(* CODESYS project beveling.project

Project tree, tasks and I/O mapping:
  Device : AM523-0808TN, Shenzhen Inovance Control Technology, version 3.5.11.50
      settings: PersistentStartAdddr = 0; PersistentStartEndAddr = 524287; Mode = 1
    application Application
      libraries: Standard, * (System); CmpEventMgr, 3.5.8.0 (System); Component Manager, 3.5.9.0 (System); CmpApp, 3.5.11.0 (System); CmpIecTask, 3.5.9.0 (System)
      task MainTask (cyclic, interval 4 ms, priority 1) calls nothing
      task ETHERCAT1 (cyclic, interval 2000 µs, priority 0) calls ETHERCAT1.EtherCAT_Task, PLC_PRG
      90_Legacy/
        program PRG_AxisDemo [ST]
      00_Types/
        data type ST_DeviceConfig
        data type ST_DeviceStatus
        data type E_AutoStep
        data type ST_ManualCommand
        data type ST_SimulationSettings
        data type ST_Recipe
        data type ST_DeviceCommand
        data type E_DeviceAction
        data type E_MachineState
        data type ST_OperatorCommand
        data type E_MachineMode
        data type ST_MachineStatus
        data type E_DeviceKind
      01_Data/
        global variables GVL_Simulation
        global variables GVL_Interface
        global variables GVL_IO
        global variables GVL_Modbus
        global variables GVL_Parameters
        global variables GVL_DeviceIds
      05_Communication/
        function block FB_ModbusInterface [ST]
      06_Simulation/
        function block FB_SimDevice [ST]
        function block FB_SimPlant [ST]
      global variables GVL_Motion
      DifferentialMonitor
      03_Units/
        function block FB_ResetLength [ST]
        function block FB_Unload [ST]
        function block FB_ClearLength [ST]
        function block FB_Initialize [ST]
        function block FB_ClearanceUnit [ST]
        function block FB_ReturnKnife [ST]
        function block FB_ClearTransfer [ST]
        function block FB_PostCut [ST]
      04_Machine/
        function F_RecipeValid [ST]
        function block FB_IOMap [ST]
        function block FB_Machine [ST]
        function block FB_AutoCycle [ST]
        function block FB_Interlocks [ST]
        function block FB_AlarmManager [ST]
        function block FB_ManualControl [ST]
      02_Devices/
        function block FB_Motor [ST]
        function F_At [ST]
        function block FB_Axis [ST]
        function block FB_DeviceManager [ST]
        function F_NextID [ST]
        function F_Done [ST]
        function block FB_Valve [ST]
        function F_Command [ST]
        function block FB_Cylinder [ST]
      program PLC_PRG [ST]
      TaskEventPreStart
    HardWare Configuration
    Network Configuration
      EtherCAT Config
      LocalBus Config
    Resources List
    ConfigStorage
    Device Diagnosis
    HwConfiguratioinDevice : SystemConfig, Inovance, version 00.00.00.10
        settings: NetworkConfigArray.NetworkConfigArray.BusType = 10; NetworkConfigArray.NetworkConfigArray.RackSum = 1; NetworkConfigArray.NetworkConfigArray.HardwareConfigArray.HardwareConfigArray.RackNo = 1
    EXP_A : 扩展卡, 汇川技术股份有限公司, version 00.00.00.10
    ETHERCAT1 : EtherCAT Master SoftMotion, 3S - Smart Software Solutions GmbH, version 3.5.11.10
        settings:  = 0; MasterCycleTime = 2000; NetworkName = 'eth1'; SelectNetworkByName = TRUE; DisableTaskGeneration = True; SlaveArrayName = ADR(_EC1_Node)
      InoSV660N : SV660_1Axis_00915, Inovance, order no. InoSV660N, version Revision=16#00010000
          settings: Number of Outputs = 6; Number of Inputs = 10; Number of Infos about Outputs = 6; Number of Infos about Inputs = 10; Configuration address of the slave = 1; Sync.Length = 18; Sync.Length = 32; FMMU.Length = 18; FMMU.Length = 32; DC sync0 cycletime = 2000; DC sync1 cycletime = 2000; Number of SDO = 10; Homing method.Index = 16#6098; Homing method.Subindex = 16#00; Homing method.Value = 1; Homing method.Size = 8; Homing method.AbortIfError = FALSE; Homing method.JumpToLine = FALSE; Homing method.Line = 0; Homing method.CompleteAccess = FALSE; Actual Position Calculation Method.Index = 16#60E6; Actual Position Calculation Method.Subindex = 16#00; Actual Position Calculation Method.Value = 0; Actual Position Calculation Method.Size = 8; Actual Position Calculation Method.AbortIfError = FALSE; Actual Position Calculation Method.JumpToLine = FALSE; Actual Position Calculation Method.Line = 0; Actual Position Calculation Method.CompleteAccess = FALSE; Speed during search for switch.Index = 16#6099; Speed during search for switch.Subindex = 16#01; Speed during search for switch.Value = 1398102; Speed during search for switch.Size = 32; Speed during search for switch.AbortIfError = FALSE; Speed during search for switch.JumpToLine = FALSE; Speed during search for switch.Line = 0; Speed during search for switch.CompleteAccess = FALSE; Homing acceleration.Index = 16#609A; Homing acceleration.Subindex = 16#00; Homing acceleration.Value = 139810133; Homing acceleration.Size = 32;
            Homing acceleration.AbortIfError = FALSE; Homing acceleration.JumpToLine = FALSE; Homing acceleration.Line = 0; Homing acceleration.CompleteAccess = FALSE; Speed during search for zero.Index = 16#6099; Speed during search for zero.Subindex = 16#02; Speed during search for zero.Value = 139810; Speed during search for zero.Size = 32; Speed during search for zero.AbortIfError = FALSE; Speed during search for zero.JumpToLine = FALSE; Speed during search for zero.Line = 0; Speed during search for zero.CompleteAccess = FALSE; Time of home searching.Index = 16#2005; Time of home searching.Subindex = 16#24; Time of home searching.Value = 50000; Time of home searching.Size = 16; Time of home searching.AbortIfError = FALSE; Time of home searching.JumpToLine = FALSE; Time of home searching.Line = 0; Time of home searching.CompleteAccess = FALSE; Positive torque limit value.Index = 16#60E0; Positive torque limit value.Subindex = 16#00; Positive torque limit value.Value = 3500; Positive torque limit value.Size = 16; Positive torque limit value.AbortIfError = FALSE; Positive torque limit value.JumpToLine = FALSE; Positive torque limit value.Line = 0; Positive torque limit value.CompleteAccess = FALSE; Negative torque limit value.Index = 16#60E1; Negative torque limit value.Subindex = 16#00; Negative torque limit value.Value = 3500; Negative torque limit value.Size = 16; Negative torque limit value.AbortIfError = FALSE; Negative torque limit value.JumpToLine = FALSE; Negative torque limit value.Line = 0; Negative torque limit value.CompleteAccess = FALSE; Max profile velocity.Index = 16#607F; Max profile velocity.Subindex = 16#00; Max profile velocity.Value = 83886080; Max profile velocity.Size = 32;
            Max profile velocity.AbortIfError = FALSE; Max profile velocity.JumpToLine = FALSE; Max profile velocity.Line = 0; Max profile velocity.CompleteAccess = FALSE; RxTxPdo.NumberofEntries = 6; RxTxPdo.Sm = 2; Controlword.Index = 16#6040; Controlword.SubIndex = 0; Controlword.Size = 16; Controlword.DependOnSlot = false; Controlword.DependOnSlotGroup = false; Target position.Index = 16#607A; Target position.SubIndex = 0; Target position.Size = 32; Target position.DependOnSlot = false; Target position.DependOnSlotGroup = false; Touch probe function.Index = 16#60B8; Touch probe function.SubIndex = 0; Touch probe function.Size = 16; Touch probe function.DependOnSlot = false; Touch probe function.DependOnSlotGroup = false; Physical outputs.Index = 16#60FE; Physical outputs.SubIndex = 1; Physical outputs.Size = 32; Physical outputs.DependOnSlot = false; Physical outputs.DependOnSlotGroup = false; Target velocity.Index = 16#60FF; Target velocity.SubIndex = 0; Target velocity.Size = 32; Target velocity.DependOnSlot = false; Target velocity.DependOnSlotGroup = false; Target torque.Index = 16#6071; Target torque.SubIndex = 0; Target torque.Size = 16; Target torque.DependOnSlot = false; Target torque.DependOnSlotGroup = false; RxTxPdo.Sm = -1; RxTxPdo.NumberofEntries = 10; RxTxPdo.Sm = 3; Error code.Index = 16#603F;
            Error code.SubIndex = 0; Error code.Size = 16; Error code.DependOnSlot = false; Error code.DependOnSlotGroup = false; Statusword.Index = 16#6041; Statusword.SubIndex = 0; Statusword.Size = 16; Statusword.DependOnSlot = false; Statusword.DependOnSlotGroup = false; Position actual value.Index = 16#6064; Position actual value.SubIndex = 0; Position actual value.Size = 32; Position actual value.DependOnSlot = false; Position actual value.DependOnSlotGroup = false; Torque actual value.Index = 16#6077; Torque actual value.SubIndex = 0; Torque actual value.Size = 16; Torque actual value.DependOnSlot = false; Torque actual value.DependOnSlotGroup = false; Following error actual value.Index = 16#60F4; Following error actual value.SubIndex = 0; Following error actual value.Size = 32; Following error actual value.DependOnSlot = false; Following error actual value.DependOnSlotGroup = false; Touch probe status.Index = 16#60B9; Touch probe status.SubIndex = 0; Touch probe status.Size = 16; Touch probe status.DependOnSlot = false; Touch probe status.DependOnSlotGroup = false; Touch probe pos1 pos value.Index = 16#60BA; Touch probe pos1 pos value.SubIndex = 0; Touch probe pos1 pos value.Size = 32; Touch probe pos1 pos value.DependOnSlot = false; Touch probe pos1 pos value.DependOnSlotGroup = false; Touch probe pos2 pos value.Index = 16#60BC; Touch probe pos2 pos value.SubIndex = 0; Touch probe pos2 pos value.Size = 32; Touch probe pos2 pos value.DependOnSlot = false; Touch probe pos2 pos value.DependOnSlotGroup = false; Digital inputs.Index = 16#60FD;
            Digital inputs.SubIndex = 0; Digital inputs.Size = 32; Digital inputs.DependOnSlot = false; Digital inputs.DependOnSlotGroup = false; Velocity actual value.Index = 16#606C; Velocity actual value.SubIndex = 0; Velocity actual value.Size = 32; Velocity actual value.DependOnSlot = false; Velocity actual value.DependOnSlotGroup = false; RxTxPdo.Sm = -1; Controlword.Name = 'Controlword'; Controlword.DataType = 'UINT'; Target position.Name = 'Target position'; Target position.DataType = 'DINT'; Touch probe function.Name = 'Touch probe function'; Touch probe function.DataType = 'UINT'; Physical outputs.Name = 'Physical outputs'; Physical outputs.DataType = 'UDINT'; Target velocity.Name = 'Target velocity'; Target velocity.DataType = 'DINT'; Target torque.Name = 'Target torque'; Target torque.DataType = 'INT'; Error code.Name = 'Error code'; Error code.DataType = 'UINT'; Statusword.Name = 'Statusword'; Statusword.DataType = 'UINT'; Position actual value.Name = 'Position actual value'; Position actual value.DataType = 'DINT'; Torque actual value.Name = 'Torque actual value'; Torque actual value.DataType = 'INT'; Following error actual value.Name = 'Following error actual value'; Following error actual value.DataType = 'DINT'; Touch probe status.Name = 'Touch probe status'; Touch probe status.DataType = 'UINT'; Touch probe pos1 pos value.Name = 'Touch probe pos1 pos value'; Touch probe pos1 pos value.DataType = 'DINT'; Touch probe pos2 pos value.Name = 'Touch probe pos2 pos value'; Touch probe pos2 pos value.DataType = 'DINT'; Digital inputs.Name = 'Digital inputs'; Digital inputs.DataType = 'UDINT';
            Velocity actual value.Name = 'Velocity actual value'; Velocity actual value.DataType = 'DINT'
          unmapped channels: Controlword, Target position, Touch probe function, Physical outputs, Target velocity, Target torque, Error code, Statusword, Position actual value, Torque actual value, Following error actual value, Touch probe status, Touch probe pos1 pos value, Touch probe pos2 pos value, Digital inputs, Velocity actual value
        Axis_1 : Axis, 3S - Smart Software Solutions GmbH, order no. 0, version 4.0.0.0
            settings: wDriveID = 0; dwRatioTechUnitsDenom = 4194304; iRatioTechUnitsNum = 5; HomingMode = 10; ZeroSignal = 0; StartDirction = 1; EndDirection = 1; PosLimitMode = 0; NegLimitMode = 0; HomingVelocity = 10; HomingApproachVelocity = 2; HomingAcceleration = 100; HomingDeceleration = 100; HomingJerk = 0; HomeMaskDistance = 0; HomePositionOffset = 0; HomePushTime = 0; HomeCompensation = 0; HomeTimeout = 0; HomeCompensationVelocity = 1000; 4000 = 1; 4001 = 0; 4003 = true; 4004 = 3; 4005 = 0; 4006 = 1.666667; 4007 = 166.666666; 4008 = 0.166667; 4009 = 50000; 4010 = 3500; 4011 = 3500; 4012 = 100.000000; ScalingIncs = 16#800000; 6005 = 10; AdrOffset_8010 = 4; BitOffset_8010 = 0; BitLength_8010 = 16; Address_8010 = '%QW2'; Type_8010 = 'UINT'; AddressPointer_8010 = ADR(%QW2);
              AdrOffset_8020 = 8; BitOffset_8020 = 0; BitLength_8020 = 32; Address_8020 = '%QD2'; Type_8020 = 'DINT'; AddressPointer_8020 = ADR(%QD2); AdrOffset_8030 = 20; BitOffset_8030 = 0; BitLength_8030 = 32; Address_8030 = '%QD5'; Type_8030 = 'DINT'; AddressPointer_8030 = ADR(%QD5); AdrOffset_8040 = 24; BitOffset_8040 = 0; BitLength_8040 = 16; Address_8040 = '%QW12'; Type_8040 = 'INT'; AddressPointer_8040 = ADR(%QW12); AdrOffset_8050 = 4294967295; BitOffset_8050 = 0; BitLength_8050 = 0; Address_8050 = ''; Type_8050 = ''; AddressPointer_8050 = 0; AdrOffset_8060 = 12; BitOffset_8060 = 0; BitLength_8060 = 16; Address_8060 = '%QW6'; Type_8060 = 'UINT'; AddressPointer_8060 = ADR(%QW6); AdrOffset_8070 = 4294967295; BitOffset_8070 = 0; BitLength_8070 = 0; Address_8070 = ''; Type_8070 = ''; AddressPointer_8070 = 0; AdrOffset_8080 = 4294967295; BitOffset_8080 = 0; BitLength_8080 = 0; Address_8080 = '';
              Type_8080 = ''; AddressPointer_8080 = 0; AdrOffset_8090 = 16; BitOffset_8090 = 0; BitLength_8090 = 32; Address_8090 = '%QD4'; Type_8090 = 'UDINT'; AddressPointer_8090 = ADR(%QD4); AdrOffset_8100 = 4294967295; BitOffset_8100 = 0; BitLength_8100 = 0; Address_8100 = ''; Type_8100 = ''; AddressPointer_8100 = 0; AdrOffset_8510 = 6; BitOffset_8510 = 0; BitLength_8510 = 16; Address_8510 = '%IW3'; Type_8510 = 'UINT'; AddressPointer_8510 = ADR(%IW3); AdrOffset_8520 = 8; BitOffset_8520 = 0; BitLength_8520 = 32; Address_8520 = '%ID2'; Type_8520 = 'DINT'; AddressPointer_8520 = ADR(%ID2); AdrOffset_8530 = 36; BitOffset_8530 = 0; BitLength_8530 = 32; Address_8530 = '%ID9'; Type_8530 = 'DINT'; AddressPointer_8530 = ADR(%ID9); AdrOffset_8540 = 12; BitOffset_8540 = 0; BitLength_8540 = 16; Address_8540 = '%IW6'; Type_8540 = 'INT'; AddressPointer_8540 = ADR(%IW6); AdrOffset_8550 = 4294967295; BitOffset_8550 = 0;
              BitLength_8550 = 0; Address_8550 = ''; Type_8550 = ''; AddressPointer_8550 = 0; AdrOffset_8560 = 32; BitOffset_8560 = 0; BitLength_8560 = 32; Address_8560 = '%ID8'; Type_8560 = 'UDINT'; AddressPointer_8560 = ADR(%ID8); AdrOffset_8570 = 20; BitOffset_8570 = 0; BitLength_8570 = 16; Address_8570 = '%IW10'; Type_8570 = 'UINT'; AddressPointer_8570 = ADR(%IW10); AdrOffset_8580 = 24; BitOffset_8580 = 0; BitLength_8580 = 32; Address_8580 = '%ID6'; Type_8580 = 'DINT'; AddressPointer_8580 = ADR(%ID6); AdrOffset_8590 = 4294967295; BitOffset_8590 = 0; BitLength_8590 = 0; Address_8590 = ''; Type_8590 = ''; AddressPointer_8590 = 0; AdrOffset_8600 = 28; BitOffset_8600 = 0; BitLength_8600 = 32; Address_8600 = '%ID7'; Type_8600 = 'DINT'; AddressPointer_8600 = ADR(%ID7); AdrOffset_8600 = 4294967295; BitOffset_8600 = 0; BitLength_8600 = 0; Address_8610 = ''; Type_8610 = ''; AddressPointer_8610 = 0;
              AdrOffset_8620 = 4; BitOffset_8620 = 0; BitLength_8620 = 16; Address_8620 = '%IW2'; Type_8620 = 'UINT'; AddressPointer_8620 = ADR(%IW2); IsValid = True; AxisNumber = 1; IsHostHoming = True; PulseSelectIndex = 4; SERVO_MAX_ID = 83886080
    SoftMotion General Axis Pool
    Serial : 串行接口, 汇川技术股份有限公司, version 00.00.00.10
      COM : Serial Port, Inovance, version 00.00.00.10
          settings: Device = AM523-0808TN; devGuid = 'e48f0cf2-85a4-455f-a8e7-135d3403221f'
    Local Bus
    EXP_B : 扩展卡, 汇川技术股份有限公司, version 00.00.00.10
    MODBUS_TCP : ModbusTCP本地从站, inovance, version 00.00.00.10
    LocalHSIO : 本地高速IO, 汇川技术股份有限公司, version 2.0.0.0
        unmapped channels: DigitalInput, DigitalOutput
    CAN : CAN总线, INOVANCE, version 00.00.00.10
*)

// Device/Application/00_Types/ST_DeviceConfig
TYPE ST_DeviceConfig :
STRUCT
eKind : E_DeviceKind;
lrInitialPosition : LREAL;
lrMinPosition : LREAL := -1000.0;
lrMaxPosition : LREAL := 1000.0;
lrMaxVelocity : LREAL := 100.0;
tSimAction : TIME := T#500MS;
END_STRUCT
END_TYPE

// Device/Application/00_Types/ST_DeviceStatus
TYPE ST_DeviceStatus :
STRUCT
xReady : BOOL;
xBusy : BOOL;
xActive : BOOL;
xError : BOOL;
udiErrorID : UDINT;
udiAcceptedID : UDINT;
udiCompletedID : UDINT;
lrPosition : LREAL;
END_STRUCT
END_TYPE

// Device/Application/00_Types/E_AutoStep
{attribute 'qualified_only'}
TYPE E_AutoStep :
(
    Idle := 0,
    FeedWait := 10,
    StopFeed := 20,
    Push := 30,
    Clearance := 40,
    Rotate := 50,
    PressDown := 60,
    KnifeDown := 70,
    SpindleOn := 80,
    Cutting := 90,
    StopCut := 100,
    PostCut := 110,
    Complete := 120,
    Fault := 900
);
END_TYPE

// Device/Application/00_Types/ST_ManualCommand
TYPE ST_ManualCommand :
STRUCT
xJogPositive : BOOL;
xJogNegative : BOOL;
xMove : BOOL;
xRun : BOOL;
lrTarget : LREAL;
lrVelocity : LREAL := 10.0;
END_STRUCT
END_TYPE

// Device/Application/00_Types/ST_SimulationSettings
TYPE ST_SimulationSettings :
STRUCT
xSafetyOK : BOOL := TRUE;
xAutoMaterial : BOOL := TRUE;
xMaterialSensor : BOOL;
tMaterialDelay : TIME := T#1S;
axStall : ARRAY[1..17] OF BOOL;
axFault : ARRAY[1..17] OF BOOL;
END_STRUCT
END_TYPE

// Device/Application/00_Types/ST_Recipe
TYPE ST_Recipe :
STRUCT
uiMaterialModel : UINT := 300;
lrCutHome : LREAL := 0.0;
lrCutLength : LREAL := 20.0;
lrCutVelocity : LREAL := 10.0;
lrPositionVelocity : LREAL := 10.0;
lrBeltVelocity : LREAL := 10.0;
lrSpindleVelocity : LREAL := 10.0;
lrLengthPosition : LREAL := 100.0;
lrLengthClear : LREAL := 0.0;
lrRotateAngle : LREAL := 0.0;
lrGripperFront : LREAL := 100.0;
lrGripperPull : LREAL := 200.0;
lrGripperBack : LREAL := 50.0;
lrGripperHome : LREAL := 0.0;
tSpray : TIME := T#300MS;
tStepTimeout : TIME := T#30S;
END_STRUCT
END_TYPE

// Device/Application/00_Types/ST_DeviceCommand
TYPE ST_DeviceCommand :
STRUCT
eAction : E_DeviceAction;
udiID : UDINT;
lrTarget : LREAL;
lrVelocity : LREAL;
END_STRUCT
END_TYPE

// Device/Application/00_Types/E_DeviceAction
{attribute 'qualified_only'}
TYPE E_DeviceAction :
(
    None := 0,
    Position := 1,
    Run := 2,
    Jog := 3,
    Stop := 4
);
END_TYPE

// Device/Application/00_Types/E_MachineState
{attribute 'qualified_only'}
TYPE E_MachineState :
(
    Stopped := 0,
    Initializing := 10,
    Ready := 20,
    Manual := 30,
    Automatic := 40,
    Fault := 90
);
END_TYPE

// Device/Application/00_Types/ST_OperatorCommand
TYPE ST_OperatorCommand :
STRUCT
eMode : E_MachineMode := E_MachineMode.Manual;
xInitialize : BOOL;
xStart : BOOL;
xStop : BOOL;
xResetAlarm : BOOL;
xContinuous : BOOL;
xRemoteControl : BOOL;
END_STRUCT
END_TYPE

// Device/Application/00_Types/E_MachineMode
{attribute 'qualified_only'}
TYPE E_MachineMode :
(
    Manual := 0,
    Automatic := 1
);
END_TYPE

// Device/Application/00_Types/ST_MachineStatus
TYPE ST_MachineStatus :
STRUCT
eState : E_MachineState;
eMode : E_MachineMode;
eAutoStep : E_AutoStep;
xSimulation : BOOL;
xRealBackendAvailable : BOOL;
xInitialized : BOOL;
xReady : BOOL;
xMaterialAtLength : BOOL;
xCycleComplete : BOOL;
udiCycleCount : UDINT;
udiAlarm : UDINT;
uiBlockedDevice : UINT;
uiManualReject : UINT;
uiClearLengthStep : UINT;
uiClearTransferStep : UINT;
uiPostStep : UINT;
uiReturnKnifeStep : UINT;
uiUnloadStep : UINT;
uiResetLengthStep : UINT;
uiInitializeStep : UINT;
uiActiveMaterialModel : UINT;
wRemoteAckSequence : WORD;
uiRemoteResult : UINT;
END_STRUCT
END_TYPE

// Device/Application/00_Types/E_DeviceKind
{attribute 'qualified_only'}
TYPE E_DeviceKind :
(
    Unused := 0,
    Axis := 1,
    Motor := 2,
    Cylinder := 3,
    Valve := 4
);
END_TYPE

// Device/Application/01_Data/GVL_Simulation
VAR_GLOBAL
    stSettings : ST_SimulationSettings;
END_VAR

// Device/Application/01_Data/GVL_Interface
VAR_GLOBAL
    stPanel : ST_OperatorCommand;
    aManual : ARRAY[1..17] OF ST_ManualCommand;
    stStatus : ST_MachineStatus;
    aDeviceStatus : ARRAY[1..17] OF ST_DeviceStatus;
END_VAR

// Device/Application/01_Data/GVL_IO
VAR_GLOBAL
    (* Unmapped interface. No AT %Q / %I bindings in this framework. *)
    xSafetyOK : BOOL;
    xMaterialAtLength : BOOL;
    axDigitalInputs : ARRAY[0..31] OF BOOL;
    axDigitalOutputs : ARRAY[0..31] OF BOOL;
    axG2RelayDemand : ARRAY[1..3] OF BOOL;
END_VAR

// Device/Application/01_Data/GVL_Modbus
VAR_GLOBAL
    (* Buffers only; the existing MODBUS_TCP driver is not bound yet. *)
    xEnable : BOOL;
    awRx : ARRAY[0..31] OF WORD;
    awTx : ARRAY[0..127] OF WORD;
END_VAR

// Device/Application/GVL_Motion
VAR_GLOBAL
    (* ================= Commands (HMI / online write) ================= *)
    xEnable     : BOOL;              (* power on / off the servo axis *)
    xReset      : BOOL;              (* reset axis error *)
    xStop       : BOOL;              (* stop and lock the axis *)
    xJogFwd     : BOOL;              (* jog forward (level) *)
    xJogRev     : BOOL;              (* jog reverse (level) *)
    xMoveRel    : BOOL;              (* relative move command (level) *)
    xMoveAbs    : BOOL;              (* absolute move command (level) *)
    xStartCycle : BOOL;              (* start auto fwd/back cycle (rising edge) *)

    rRelDist    : LREAL := 100.0;    (* relative move distance [mm] *)
    rTargetPos  : LREAL := 0.0;      (* absolute target position [mm] *)

    (* ================= Motion parameters ================= *)
    rJogVel     : LREAL := 10.0;     (* jog velocity [mm/s] *)
    rVel        : LREAL := 30.0;     (* positioning velocity [mm/s] *)
    rAcc        : LREAL := 200.0;    (* acceleration [mm/s2] *)
    rDec        : LREAL := 200.0;    (* deceleration [mm/s2] *)
    rStroke     : LREAL := 100.0;    (* auto cycle stroke (one way) [mm] *)
    tDwell      : TIME  := T#1S;     (* dwell time at cycle ends *)

    (* ================= Status ================= *)
    xPowered    : BOOL;              (* MC_Power.Status : servo enabled *)
    xAxisReady  : BOOL;              (* axis in StandStill -> motion allowed *)
    xBusy       : BOOL;              (* any motion active *)
    xDisabled   : BOOL;              (* axis state = Disabled *)
    xStandStill : BOOL;              (* axis state = StandStill *)
    xStopping   : BOOL;              (* axis state = Stopping *)
    xErrorStop  : BOOL;              (* axis state = ErrorStop *)
    xAxisError  : BOOL;              (* axis reports an error *)
    iAxisErrorID: DWORD;             (* axis error code *)
    rActPos     : LREAL;             (* actual position [mm] *)
    iState      : INT;               (* auto cycle step number *)
END_VAR

// Device/Application/01_Data/GVL_Parameters
VAR_GLOBAL
    (* Simulation examples only: these are NOT commissioned machine settings. *)
    xSimulation : BOOL := TRUE;
    stRecipe : ST_Recipe;
END_VAR

// Device/Application/01_Data/GVL_DeviceIds
VAR_GLOBAL CONSTANT
    D1_Belt : UINT := 1;
    D2_CutFeed : UINT := 2;
    D3_Spindle : UINT := 3;
    D4_LengthMove : UINT := 4;
    D5_LengthLift : UINT := 5;
    D7_GripperMove : UINT := 7;
    D8_Rotate : UINT := 8;
    G1_Press : UINT := 9;
    G2_SideStop : UINT := 10;
    G3_Push : UINT := 11;
    G4_RollerLift : UINT := 12;
    G5_Spray : UINT := 13;
    G6_Air : UINT := 14;
    G7_GripperLift : UINT := 15;
    G8_GripperClamp : UINT := 16;
    G9_KnifeLift : UINT := 17;
END_VAR

// Device/Application/PLC_PRG
PROGRAM PLC_PRG
VAR
    fbCommunication : FB_ModbusInterface;
    fbMachine : FB_Machine;
    fbIO : FB_IOMap;
END_VAR

(* One cyclic owner in ETHERCAT1. All lower device FBs are called each scan. *)
fbCommunication(xEnable:=GVL_Modbus.xEnable,stStatus:=GVL_Interface.stStatus,
    aStatus:=GVL_Interface.aDeviceStatus,awRx:=GVL_Modbus.awRx,awTx:=GVL_Modbus.awTx);
fbMachine(xSimulation:=GVL_Parameters.xSimulation,stPanel:=GVL_Interface.stPanel,
    stRemote:=fbCommunication.stCommand,xRemoteRequest:=fbCommunication.xRequest,
    wRemoteSequence:=fbCommunication.wRequestSequence,aManual:=GVL_Interface.aManual,
    stRecipe:=GVL_Parameters.stRecipe,stSim:=GVL_Simulation.stSettings,
    xRealSafetyOK:=GVL_IO.xSafetyOK,xRealMaterial:=GVL_IO.xMaterialAtLength);
GVL_Interface.stStatus:=fbMachine.stStatus;
GVL_Interface.aDeviceStatus:=fbMachine.aDeviceStatus;
fbIO(uiMaterialModel:=fbMachine.stStatus.uiActiveMaterialModel,aCommand:=fbMachine.aSelectedCommand,
    aStatus:=fbMachine.aDeviceStatus,
    axOutputs:=GVL_IO.axDigitalOutputs,axG2RelayDemand:=GVL_IO.axG2RelayDemand);

END_PROGRAM

// Device/Application/05_Communication/FB_ModbusInterface
FUNCTION_BLOCK FB_ModbusInterface
VAR_INPUT
    xEnable : BOOL;
    stStatus : ST_MachineStatus;
    aStatus : ARRAY[1..17] OF ST_DeviceStatus;
END_VAR
VAR_IN_OUT
    awRx : ARRAY[0..31] OF WORD;
    awTx : ARRAY[0..127] OF WORD;
END_VAR
VAR_OUTPUT
    xRequest : BOOL;
    wRequestSequence : WORD;
    stCommand : ST_OperatorCommand;
    uiParseResult : UINT;
END_VAR
VAR
    aSnapshot : ARRAY[0..31] OF WORD;
    wLastSeen : WORD;
    xWasEnabled : BOOL;
    i : INT;
END_VAR

xRequest:=FALSE;
stCommand.xInitialize:=FALSE; stCommand.xStart:=FALSE;
stCommand.xStop:=FALSE; stCommand.xResetAlarm:=FALSE;
IF NOT xEnable OR NOT xWasEnabled THEN
    (* Baseline on enable, so reconnect never replays a stale command. *)
    wLastSeen:=awRx[1];
ELSIF (awRx[1]<>0) AND (awRx[1]<>wLastSeen) THEN
    aSnapshot:=awRx;
    IF aSnapshot[1]=awRx[1] THEN
        wLastSeen:=aSnapshot[1]; wRequestSequence:=aSnapshot[1]; uiParseResult:=0;
        IF (aSnapshot[0]<>1) OR (aSnapshot[3]>1) OR (aSnapshot[2]<1) OR (aSnapshot[2]>4) THEN
            uiParseResult:=2;
        ELSE
            IF aSnapshot[3]=0 THEN stCommand.eMode:=E_MachineMode.Manual;
            ELSE stCommand.eMode:=E_MachineMode.Automatic; END_IF
            stCommand.xContinuous:=aSnapshot[4]<>0;
            CASE aSnapshot[2] OF
            1: stCommand.xInitialize:=TRUE;
            2: stCommand.xStart:=TRUE;
            3: stCommand.xStop:=TRUE;
            4: stCommand.xResetAlarm:=TRUE;
            END_CASE
            xRequest:=TRUE;
        END_IF
    END_IF
END_IF
xWasEnabled:=xEnable;
FOR i:=0 TO 127 DO awTx[i]:=0; END_FOR
awTx[0]:=1; awTx[1]:=stStatus.wRemoteAckSequence; awTx[2]:=UINT_TO_WORD(stStatus.uiRemoteResult);
awTx[3]:=TO_WORD(stStatus.eState); awTx[4]:=TO_WORD(stStatus.eAutoStep);
awTx[5]:=UDINT_TO_WORD(stStatus.udiAlarm); awTx[6]:=UDINT_TO_WORD(SHR(stStatus.udiAlarm,16));
awTx[7]:=UDINT_TO_WORD(stStatus.udiCycleCount); awTx[8]:=UDINT_TO_WORD(SHR(stStatus.udiCycleCount,16));
awTx[9]:=BOOL_TO_WORD(stStatus.xSimulation); awTx[10]:=BOOL_TO_WORD(stStatus.xInitialized);
awTx[11]:=BOOL_TO_WORD(stStatus.xMaterialAtLength); awTx[12]:=UINT_TO_WORD(stStatus.uiActiveMaterialModel);
awTx[13]:=wRequestSequence; awTx[14]:=UINT_TO_WORD(uiParseResult);
(* Positions at [32..48]: signed INT, 0.1 engineering-unit scaling. *)
FOR i:=1 TO 17 DO awTx[31+i]:=INT_TO_WORD(LREAL_TO_INT(aStatus[i].lrPosition*10.0)); END_FOR

END_FUNCTION_BLOCK

// Device/Application/04_Machine/FB_Machine
FUNCTION_BLOCK FB_Machine
VAR_INPUT
    xSimulation : BOOL;
    stPanel : ST_OperatorCommand;
    stRemote : ST_OperatorCommand;
    xRemoteRequest : BOOL;
    wRemoteSequence : WORD;
    aManual : ARRAY[1..17] OF ST_ManualCommand;
    stRecipe : ST_Recipe;
    stSim : ST_SimulationSettings;
    xRealSafetyOK : BOOL;
    xRealMaterial : BOOL;
END_VAR
VAR_OUTPUT
    stStatus : ST_MachineStatus;
    aDeviceStatus : ARRAY[1..17] OF ST_DeviceStatus;
    aSelectedCommand : ARRAY[1..17] OF ST_DeviceCommand;
END_VAR
VAR
    stCommand : ST_OperatorCommand;
    stActiveRecipe : ST_Recipe;
    aRequest : ARRAY[1..17] OF ST_DeviceCommand;
    stEmpty : ST_DeviceCommand;
    fbDevices : FB_DeviceManager;
    fbManual : FB_ManualControl;
    fbAuto : FB_AutoCycle;
    fbInitialize : FB_Initialize;
    fbInterlocks : FB_Interlocks;
    fbPlant : FB_SimPlant;
    fbAlarm : FB_AlarmManager;
    rtInitialize : R_TRIG;
    rtStart : R_TRIG;
    rtReset : R_TRIG;
    udiCounter : UDINT;
    udiFault : UDINT;
    xSafetyOK : BOOL;
    xMaterial : BOOL;
    xInitialized : BOOL;
    xPermit : BOOL;
    xRemoteAccepted : BOOL;
    xResetDevices : BOOL;
    xLastSimulation : BOOL := TRUE;
    xManualReleased : BOOL;
    xManualArmed : BOOL;
    eActiveMode : E_MachineMode;
    i : INT;
END_VAR

stCommand:=stPanel;
IF stPanel.xRemoteControl THEN
    (* Mode and continuous selection persist between remote command frames. *)
    stCommand.eMode:=stRemote.eMode;
    stCommand.xContinuous:=stRemote.xContinuous;
END_IF
xRemoteAccepted:=FALSE;
IF xRemoteRequest THEN
    stStatus.wRemoteAckSequence:=wRemoteSequence;
    IF stPanel.xRemoteControl THEN
        stCommand:=stRemote;
        (* Local stop always overrides remote control. *)
        stCommand.xStop:=stCommand.xStop OR stPanel.xStop;
        stStatus.uiRemoteResult:=0; xRemoteAccepted:=TRUE;
    ELSE stStatus.uiRemoteResult:=1;
    END_IF
END_IF
rtInitialize(CLK:=stCommand.xInitialize);
rtStart(CLK:=stCommand.xStart);
rtReset(CLK:=stCommand.xResetAlarm);
IF xSimulation THEN xSafetyOK:=stSim.xSafetyOK; xMaterial:=fbPlant.xMaterialAtLength;
ELSE xSafetyOK:=xRealSafetyOK; xMaterial:=xRealMaterial; END_IF
udiFault:=0;
IF NOT xSafetyOK THEN udiFault:=1001; END_IF
IF NOT xSimulation THEN udiFault:=3001; END_IF
IF xSimulation<>xLastSimulation THEN
    stStatus.eState:=E_MachineState.Stopped; xInitialized:=FALSE;
END_IF
xLastSimulation:=xSimulation;
FOR i:=1 TO 17 DO
    IF aDeviceStatus[i].xError THEN udiFault:=10000+INT_TO_UDINT(i); END_IF
    aRequest[i]:=stEmpty;
END_FOR
IF (stStatus.eState=E_MachineState.Automatic) OR (stStatus.eState=E_MachineState.Manual) THEN
    IF stCommand.eMode<>eActiveMode THEN stStatus.eState:=E_MachineState.Stopped; xInitialized:=FALSE; END_IF
END_IF
IF stCommand.xStop THEN stStatus.eState:=E_MachineState.Stopped; xInitialized:=FALSE; END_IF
IF udiFault<>0 THEN stStatus.eState:=E_MachineState.Fault; xInitialized:=FALSE; END_IF
xResetDevices:=rtReset.Q AND xSafetyOK AND xSimulation;
IF xResetDevices THEN
    (* Reset injected/device errors before clearing the machine latch next scan. *)
    udiFault:=0;
    FOR i:=1 TO 17 DO IF stSim.axFault[i] THEN udiFault:=10000+INT_TO_UDINT(i); END_IF END_FOR
END_IF
fbAlarm(udiIncoming:=udiFault,xReset:=xResetDevices);
IF (stStatus.eState=E_MachineState.Fault) AND (fbAlarm.udiLatched=0) AND xResetDevices THEN
    stStatus.eState:=E_MachineState.Stopped;
END_IF
IF fbAlarm.udiLatched<>0 THEN stStatus.eState:=E_MachineState.Fault; END_IF
IF rtInitialize.Q AND NOT stCommand.xStop THEN
    IF (stStatus.eState=E_MachineState.Stopped) AND xSimulation AND xSafetyOK AND F_RecipeValid(stRecipe) THEN
        stActiveRecipe:=stRecipe; stStatus.eState:=E_MachineState.Initializing;
        eActiveMode:=stCommand.eMode; xInitialized:=FALSE;
    ELSIF xRemoteAccepted THEN stStatus.uiRemoteResult:=3;
    END_IF
END_IF
IF stStatus.eState=E_MachineState.Ready THEN
    IF stCommand.eMode=E_MachineMode.Manual THEN
        stStatus.eState:=E_MachineState.Manual; eActiveMode:=E_MachineMode.Manual;
    ELSIF rtStart.Q AND NOT stCommand.xStop THEN
        IF F_RecipeValid(stRecipe) THEN
            stActiveRecipe:=stRecipe; eActiveMode:=E_MachineMode.Automatic;
            stStatus.eState:=E_MachineState.Automatic;
        ELSIF xRemoteAccepted THEN stStatus.uiRemoteResult:=5;
        END_IF
    END_IF
ELSIF (stStatus.eState=E_MachineState.Manual) AND (stCommand.eMode=E_MachineMode.Automatic) THEN
    stStatus.eState:=E_MachineState.Stopped; xInitialized:=FALSE;
END_IF
IF rtStart.Q AND xRemoteAccepted AND (stStatus.eState<>E_MachineState.Automatic) THEN stStatus.uiRemoteResult:=3; END_IF

xManualReleased:=TRUE;
FOR i:=1 TO 17 DO
    IF aManual[i].xJogPositive OR aManual[i].xJogNegative OR aManual[i].xMove OR aManual[i].xRun THEN xManualReleased:=FALSE; END_IF
END_FOR
IF stStatus.eState<>E_MachineState.Manual THEN xManualArmed:=FALSE;
ELSIF xManualReleased THEN xManualArmed:=TRUE;
END_IF
fbInitialize(xExecute:=stStatus.eState=E_MachineState.Initializing,stRecipe:=stActiveRecipe,
    aCommand:=aRequest,aStatus:=aDeviceStatus,udiCounter:=udiCounter);
fbManual(xEnable:=(stStatus.eState=E_MachineState.Manual) AND xManualArmed,
    aManual:=aManual,aCommand:=aRequest,aStatus:=aDeviceStatus,udiCounter:=udiCounter);
fbAuto(xRun:=stStatus.eState=E_MachineState.Automatic,xContinuous:=stCommand.xContinuous,
    xMaterialAtLength:=xMaterial,stRecipe:=stActiveRecipe,aCommand:=aRequest,aStatus:=aDeviceStatus,udiCounter:=udiCounter);
IF fbInitialize.xDone THEN xInitialized:=TRUE; stStatus.eState:=E_MachineState.Ready; END_IF
IF fbInitialize.xError OR fbAuto.xError THEN
    udiFault:=MAX(fbInitialize.udiErrorID,fbAuto.udiErrorID);
    fbAlarm(udiIncoming:=udiFault,xReset:=FALSE);
    stStatus.eState:=E_MachineState.Fault; xInitialized:=FALSE;
END_IF
IF fbAuto.xDone THEN
    stStatus.udiCycleCount:=stStatus.udiCycleCount+1;
    IF NOT stCommand.xContinuous THEN stStatus.eState:=E_MachineState.Ready; END_IF
END_IF
xPermit:=xSimulation AND xSafetyOK AND NOT stCommand.xStop AND (fbAlarm.udiLatched=0)
    AND ((stStatus.eState=E_MachineState.Initializing) OR (stStatus.eState=E_MachineState.Manual)
    OR (stStatus.eState=E_MachineState.Automatic));
fbInterlocks(xPermit:=xPermit,stRecipe:=stActiveRecipe,aRequest:=aRequest,aStatus:=aDeviceStatus);
aSelectedCommand:=fbInterlocks.aCommand;
fbDevices(xEnable:=xSimulation AND xSafetyOK,xSimulation:=xSimulation,xReset:=xResetDevices,
    stSim:=stSim,aCommand:=aSelectedCommand);
aDeviceStatus:=fbDevices.aStatus;
fbPlant(xEnable:=xSimulation,stSettings:=stSim,aStatus:=aDeviceStatus);
stStatus.eMode:=stCommand.eMode; stStatus.eAutoStep:=fbAuto.eStep;
stStatus.xSimulation:=xSimulation; stStatus.xRealBackendAvailable:=FALSE;
stStatus.xInitialized:=xInitialized;
stStatus.xReady:=xInitialized AND (stStatus.eState=E_MachineState.Ready);
stStatus.xMaterialAtLength:=xMaterial; stStatus.xCycleComplete:=fbAuto.xDone;
stStatus.udiAlarm:=fbAlarm.udiLatched; stStatus.uiBlockedDevice:=fbInterlocks.uiBlockedDevice;
stStatus.uiManualReject:=fbManual.uiRejectDevice;
stStatus.uiClearLengthStep:=fbAuto.uiClearLengthStep; stStatus.uiClearTransferStep:=fbAuto.uiClearTransferStep;
stStatus.uiPostStep:=fbAuto.uiPostStep; stStatus.uiReturnKnifeStep:=fbAuto.uiReturnKnifeStep;
stStatus.uiUnloadStep:=fbAuto.uiUnloadStep; stStatus.uiResetLengthStep:=fbAuto.uiResetLengthStep;
stStatus.uiInitializeStep:=fbInitialize.uiStep; stStatus.uiActiveMaterialModel:=stActiveRecipe.uiMaterialModel;

END_FUNCTION_BLOCK

// Device/Application/04_Machine/F_RecipeValid
FUNCTION F_RecipeValid : BOOL
VAR_INPUT
    stRecipe : ST_Recipe;
END_VAR

F_RecipeValid := ((stRecipe.uiMaterialModel = 300) OR
    (stRecipe.uiMaterialModel = 400) OR (stRecipe.uiMaterialModel = 600))
    AND (stRecipe.lrCutLength > 0.0) AND (stRecipe.lrCutLength <= 500.0)
    AND (stRecipe.lrCutVelocity > 0.0) AND (stRecipe.lrCutVelocity <= 100.0)
    AND (stRecipe.lrPositionVelocity > 0.0) AND (stRecipe.lrPositionVelocity <= 100.0)
    AND (stRecipe.lrBeltVelocity > 0.0) AND (stRecipe.lrBeltVelocity <= 100.0)
    AND (stRecipe.lrSpindleVelocity > 0.0) AND (stRecipe.lrSpindleVelocity <= 100.0)
    AND (stRecipe.tStepTimeout >= T#1S) AND (stRecipe.tSpray > T#0MS)
    AND (ABS(stRecipe.lrCutHome) <= 500.0)
    AND (ABS(stRecipe.lrCutHome + stRecipe.lrCutLength) <= 1000.0)
    AND (ABS(stRecipe.lrLengthPosition) <= 1000.0)
    AND (ABS(stRecipe.lrLengthClear) <= 1000.0)
    AND (ABS(stRecipe.lrRotateAngle) <= 360.0)
    AND (stRecipe.lrGripperHome < stRecipe.lrGripperBack)
    AND (stRecipe.lrGripperBack < stRecipe.lrGripperFront)
    AND (stRecipe.lrGripperFront < stRecipe.lrGripperPull)
    AND (ABS(stRecipe.lrGripperPull) <= 1000.0);

END_FUNCTION

// Device/Application/02_Devices/FB_DeviceManager
FUNCTION_BLOCK FB_DeviceManager
VAR_INPUT
    xEnable : BOOL;
    xSimulation : BOOL;
    xReset : BOOL;
    stSim : ST_SimulationSettings;
    aCommand : ARRAY[1..17] OF ST_DeviceCommand;
END_VAR
VAR_OUTPUT
    aStatus : ARRAY[1..17] OF ST_DeviceStatus;
END_VAR
VAR
    aConfig : ARRAY[1..17] OF ST_DeviceConfig;
    aAxis : ARRAY[1..17] OF FB_Axis;
    aMotor : ARRAY[1..17] OF FB_Motor;
    aCylinder : ARRAY[1..17] OF FB_Cylinder;
    aValve : ARRAY[1..17] OF FB_Valve;
    xBooted : BOOL;
    i : INT;
END_VAR

IF NOT xBooted THEN
    aConfig[1].eKind := E_DeviceKind.Motor;
    aConfig[2].eKind := E_DeviceKind.Axis;
    aConfig[3].eKind := E_DeviceKind.Motor;
    aConfig[4].eKind := E_DeviceKind.Axis;
    (* D5 is modeled as a positioning lift; 0/1 are simulation up/down points. *)
    aConfig[5].eKind := E_DeviceKind.Axis;
    aConfig[7].eKind := E_DeviceKind.Axis;
    aConfig[8].eKind := E_DeviceKind.Axis;
    FOR i := 9 TO 17 DO aConfig[i].eKind := E_DeviceKind.Cylinder; END_FOR
    aConfig[13].eKind := E_DeviceKind.Valve;
    aConfig[14].eKind := E_DeviceKind.Valve;
    aConfig[12].lrInitialPosition := 1.0;
    FOR i := 1 TO 17 DO
        IF aConfig[i].eKind = E_DeviceKind.Cylinder THEN
            aConfig[i].lrMinPosition := 0.0; aConfig[i].lrMaxPosition := 1.0;
        END_IF
    END_FOR
    xBooted := TRUE;
END_IF
FOR i := 1 TO 17 DO
    CASE aConfig[i].eKind OF
    E_DeviceKind.Axis:
        aAxis[i](xSimulation:=xSimulation,xEnable:=xEnable,xReset:=xReset,
            xStall:=stSim.axStall[i],xInjectFault:=stSim.axFault[i],stConfig:=aConfig[i],stCommand:=aCommand[i]);
        aStatus[i] := aAxis[i].stStatus;
    E_DeviceKind.Motor:
        aMotor[i](xSimulation:=xSimulation,xEnable:=xEnable,xReset:=xReset,
            xStall:=stSim.axStall[i],xInjectFault:=stSim.axFault[i],stConfig:=aConfig[i],stCommand:=aCommand[i]);
        aStatus[i] := aMotor[i].stStatus;
    E_DeviceKind.Cylinder:
        aCylinder[i](xSimulation:=xSimulation,xEnable:=xEnable,xReset:=xReset,
            xStall:=stSim.axStall[i],xInjectFault:=stSim.axFault[i],stConfig:=aConfig[i],stCommand:=aCommand[i]);
        aStatus[i] := aCylinder[i].stStatus;
    E_DeviceKind.Valve:
        aValve[i](xSimulation:=xSimulation,xEnable:=xEnable,xReset:=xReset,
            xStall:=stSim.axStall[i],xInjectFault:=stSim.axFault[i],stConfig:=aConfig[i],stCommand:=aCommand[i]);
        aStatus[i] := aValve[i].stStatus;
    END_CASE
END_FOR

END_FUNCTION_BLOCK

// Device/Application/02_Devices/FB_Axis
FUNCTION_BLOCK FB_Axis
VAR_INPUT
    xSimulation : BOOL;
    xEnable : BOOL;
    xReset : BOOL;
    xStall : BOOL;
    xInjectFault : BOOL;
    stConfig : ST_DeviceConfig;
    stCommand : ST_DeviceCommand;
END_VAR
VAR_OUTPUT
    stStatus : ST_DeviceStatus;
END_VAR
VAR
    fbSimulation : FB_SimDevice;
END_VAR

(* The real hardware adapter is intentionally not commissioned. *)
fbSimulation(xEnable := xEnable AND xSimulation, xReset := xReset,
    xStall := xStall, xInjectFault := xInjectFault,
    stConfig := stConfig, stCommand := stCommand);
stStatus := fbSimulation.stStatus;
IF NOT xSimulation THEN
    stStatus.xReady := FALSE; stStatus.xBusy := FALSE; stStatus.xActive := FALSE;
    stStatus.xError := TRUE; stStatus.udiErrorID := 3001;
END_IF

END_FUNCTION_BLOCK

// Device/Application/06_Simulation/FB_SimDevice
FUNCTION_BLOCK FB_SimDevice
VAR_INPUT
    xEnable : BOOL;
    xReset : BOOL;
    xStall : BOOL;
    xInjectFault : BOOL;
    stConfig : ST_DeviceConfig;
    stCommand : ST_DeviceCommand;
END_VAR
VAR_OUTPUT
    stStatus : ST_DeviceStatus;
END_VAR
VAR
    xBooted : BOOL;
    xAction : BOOL;
    udiLastID : UDINT;
    lrStart : LREAL;
    lrTarget : LREAL;
    lrJogDelta : LREAL;
    tLastJog : TIME;
    tonAction : TON;
    tonJog : TON;
END_VAR

IF NOT xBooted THEN
    stStatus.lrPosition := stConfig.lrInitialPosition;
    xBooted := TRUE;
END_IF
IF xReset AND NOT xInjectFault THEN
    stStatus.xError := FALSE; stStatus.udiErrorID := 0;
END_IF
IF xInjectFault THEN stStatus.xError := TRUE; stStatus.udiErrorID := 9001; END_IF
stStatus.xReady := xEnable AND NOT stStatus.xError AND (stConfig.eKind <> E_DeviceKind.Unused);

IF NOT stStatus.xReady OR (stCommand.eAction = E_DeviceAction.None)
   OR (stCommand.eAction = E_DeviceAction.Stop) THEN
    xAction := FALSE; udiLastID := 0;
    stStatus.xBusy := FALSE; stStatus.xActive := FALSE;
    stStatus.udiAcceptedID := 0; stStatus.udiCompletedID := 0;
ELSIF (stCommand.udiID <> 0) AND (stCommand.udiID <> udiLastID) THEN
    udiLastID := stCommand.udiID;
    stStatus.udiAcceptedID := udiLastID; stStatus.udiCompletedID := 0;
    lrStart := stStatus.lrPosition; lrTarget := stCommand.lrTarget;
    IF (ABS(stCommand.lrVelocity) > stConfig.lrMaxVelocity)
       OR ((stCommand.eAction = E_DeviceAction.Position) AND
           ((lrTarget < stConfig.lrMinPosition) OR (lrTarget > stConfig.lrMaxPosition))) THEN
        stStatus.xError := TRUE; stStatus.udiErrorID := 2001; xAction := FALSE;
    ELSE
        xAction := stCommand.eAction <> E_DeviceAction.Jog;
        stStatus.xBusy := TRUE; stStatus.xActive := FALSE;
    END_IF
    (* Reset on acceptance; the regular call below starts the new timer. *)
    tonAction(IN := FALSE);
END_IF
tonAction(IN := xAction AND stStatus.xReady, PT := stConfig.tSimAction);
IF xAction AND NOT xStall AND stStatus.xReady THEN
    IF stCommand.eAction = E_DeviceAction.Position THEN
        stStatus.lrPosition := lrStart + (lrTarget-lrStart) *
            MIN(1.0, TIME_TO_LREAL(tonAction.ET) / MAX(1.0, TIME_TO_LREAL(stConfig.tSimAction)));
    END_IF
    IF tonAction.Q THEN
        IF stCommand.eAction = E_DeviceAction.Position THEN stStatus.lrPosition := lrTarget; END_IF
        stStatus.xBusy := FALSE;
        stStatus.xActive := stCommand.eAction = E_DeviceAction.Run;
        stStatus.udiCompletedID := udiLastID;
        xAction := FALSE;
    END_IF
END_IF
tonJog(IN := stStatus.xReady AND (stCommand.eAction = E_DeviceAction.Jog), PT := T#24H);
IF tonJog.IN THEN
    lrJogDelta := TIME_TO_LREAL(tonJog.ET-tLastJog) / 1000.0;
    IF NOT xStall THEN
        stStatus.lrPosition := LIMIT(stConfig.lrMinPosition,
            stStatus.lrPosition+stCommand.lrVelocity*lrJogDelta, stConfig.lrMaxPosition);
    END_IF
    stStatus.xBusy := TRUE; stStatus.xActive := TRUE;
    tLastJog := tonJog.ET;
ELSE tLastJog := T#0MS;
END_IF
IF stStatus.xError THEN
    stStatus.xReady := FALSE; stStatus.xBusy := FALSE; stStatus.xActive := FALSE;
END_IF

END_FUNCTION_BLOCK

// Device/Application/02_Devices/FB_Motor
FUNCTION_BLOCK FB_Motor
VAR_INPUT
    xSimulation : BOOL;
    xEnable : BOOL;
    xReset : BOOL;
    xStall : BOOL;
    xInjectFault : BOOL;
    stConfig : ST_DeviceConfig;
    stCommand : ST_DeviceCommand;
END_VAR
VAR_OUTPUT
    stStatus : ST_DeviceStatus;
END_VAR
VAR
    fbSimulation : FB_SimDevice;
END_VAR

(* The real hardware adapter is intentionally not commissioned. *)
fbSimulation(xEnable := xEnable AND xSimulation, xReset := xReset,
    xStall := xStall, xInjectFault := xInjectFault,
    stConfig := stConfig, stCommand := stCommand);
stStatus := fbSimulation.stStatus;
IF NOT xSimulation THEN
    stStatus.xReady := FALSE; stStatus.xBusy := FALSE; stStatus.xActive := FALSE;
    stStatus.xError := TRUE; stStatus.udiErrorID := 3001;
END_IF

END_FUNCTION_BLOCK

// Device/Application/02_Devices/FB_Cylinder
FUNCTION_BLOCK FB_Cylinder
VAR_INPUT
    xSimulation : BOOL;
    xEnable : BOOL;
    xReset : BOOL;
    xStall : BOOL;
    xInjectFault : BOOL;
    stConfig : ST_DeviceConfig;
    stCommand : ST_DeviceCommand;
END_VAR
VAR_OUTPUT
    stStatus : ST_DeviceStatus;
END_VAR
VAR
    fbSimulation : FB_SimDevice;
END_VAR

(* The real hardware adapter is intentionally not commissioned. *)
fbSimulation(xEnable := xEnable AND xSimulation, xReset := xReset,
    xStall := xStall, xInjectFault := xInjectFault,
    stConfig := stConfig, stCommand := stCommand);
stStatus := fbSimulation.stStatus;
IF NOT xSimulation THEN
    stStatus.xReady := FALSE; stStatus.xBusy := FALSE; stStatus.xActive := FALSE;
    stStatus.xError := TRUE; stStatus.udiErrorID := 3001;
END_IF

END_FUNCTION_BLOCK

// Device/Application/02_Devices/FB_Valve
FUNCTION_BLOCK FB_Valve
VAR_INPUT
    xSimulation : BOOL;
    xEnable : BOOL;
    xReset : BOOL;
    xStall : BOOL;
    xInjectFault : BOOL;
    stConfig : ST_DeviceConfig;
    stCommand : ST_DeviceCommand;
END_VAR
VAR_OUTPUT
    stStatus : ST_DeviceStatus;
END_VAR
VAR
    fbSimulation : FB_SimDevice;
END_VAR

(* The real hardware adapter is intentionally not commissioned. *)
fbSimulation(xEnable := xEnable AND xSimulation, xReset := xReset,
    xStall := xStall, xInjectFault := xInjectFault,
    stConfig := stConfig, stCommand := stCommand);
stStatus := fbSimulation.stStatus;
IF NOT xSimulation THEN
    stStatus.xReady := FALSE; stStatus.xBusy := FALSE; stStatus.xActive := FALSE;
    stStatus.xError := TRUE; stStatus.udiErrorID := 3001;
END_IF

END_FUNCTION_BLOCK

// Device/Application/04_Machine/FB_ManualControl
FUNCTION_BLOCK FB_ManualControl
VAR_INPUT
    xEnable : BOOL;
    aManual : ARRAY[1..17] OF ST_ManualCommand;
END_VAR
VAR_IN_OUT
    aCommand : ARRAY[1..17] OF ST_DeviceCommand;
    aStatus : ARRAY[1..17] OF ST_DeviceStatus;
    udiCounter : UDINT;
END_VAR
VAR_OUTPUT
    uiRejectDevice : UINT;
END_VAR
VAR
    aPrev : ARRAY[1..17] OF ST_ManualCommand;
    aPending : ARRAY[1..17] OF ST_DeviceCommand;
    aRunID : ARRAY[1..17] OF UDINT;
    i : INT;
    lrVelocity : LREAL;
END_VAR

uiRejectDevice:=0;
FOR i:=1 TO 17 DO
    IF NOT xEnable THEN
        aPending[i].eAction:=E_DeviceAction.None;
        aRunID[i]:=0;
    ELSIF i<>6 THEN
        lrVelocity:=LIMIT(0.1,ABS(aManual[i].lrVelocity),100.0);
        IF (aManual[i].xJogPositive AND aManual[i].xJogNegative)
           OR ((aManual[i].xJogPositive OR aManual[i].xJogNegative) AND (aManual[i].xMove OR aManual[i].xRun))
           OR (aManual[i].xMove AND aManual[i].xRun) THEN
            uiRejectDevice:=INT_TO_UINT(i); aPending[i].eAction:=E_DeviceAction.None;
        ELSIF aManual[i].xJogPositive OR aManual[i].xJogNegative THEN
            aPending[i].eAction:=E_DeviceAction.None;
            IF aRunID[i]=0 THEN aRunID[i]:=F_NextID(udiCounter); END_IF
            IF aManual[i].xJogNegative THEN lrVelocity:=-lrVelocity; END_IF
            IF (i=2) OR (i=4) OR (i=5) OR (i=7) OR (i=8) THEN
                aCommand[i]:=F_Command(E_DeviceAction.Jog,aRunID[i],0.0,lrVelocity);
            ELSE uiRejectDevice:=INT_TO_UINT(i);
            END_IF
        ELSIF aManual[i].xRun THEN
            aPending[i].eAction:=E_DeviceAction.None;
            IF (i=1) OR (i=3) OR (i=13) OR (i=14) THEN
                IF aRunID[i]=0 THEN aRunID[i]:=F_NextID(udiCounter); END_IF
                aCommand[i]:=F_Command(E_DeviceAction.Run,aRunID[i],0.0,lrVelocity);
            ELSE uiRejectDevice:=INT_TO_UINT(i);
            END_IF
        ELSE
            aRunID[i]:=0;
            IF aManual[i].xMove AND NOT aPrev[i].xMove THEN
                IF (i<>1) AND (i<>3) AND (i<>13) AND (i<>14) THEN
                    aPending[i]:=F_Command(E_DeviceAction.Position,F_NextID(udiCounter),aManual[i].lrTarget,lrVelocity);
                ELSE uiRejectDevice:=INT_TO_UINT(i);
                END_IF
            END_IF
            IF aPending[i].eAction<>E_DeviceAction.None THEN
                aCommand[i]:=aPending[i];
                IF F_Done(aStatus[i],aPending[i].udiID) THEN aPending[i].eAction:=E_DeviceAction.None; END_IF
            END_IF
        END_IF
    END_IF
    (* Synchronize while disabled: held buttons never acquire a fresh move edge. *)
    aPrev[i]:=aManual[i];
END_FOR

END_FUNCTION_BLOCK

// Device/Application/02_Devices/F_NextID
FUNCTION F_NextID : UDINT
VAR_IN_OUT
    udiCounter : UDINT;
END_VAR

IF udiCounter = 16#FFFFFFFF THEN udiCounter := 1;
ELSE udiCounter := udiCounter + 1;
END_IF
F_NextID := udiCounter;

END_FUNCTION

// Device/Application/02_Devices/F_Command
FUNCTION F_Command : ST_DeviceCommand
VAR_INPUT
    eAction : E_DeviceAction;
    udiID : UDINT;
    lrTarget : LREAL;
    lrVelocity : LREAL;
END_VAR

F_Command.eAction := eAction;
F_Command.udiID := udiID;
F_Command.lrTarget := lrTarget;
F_Command.lrVelocity := lrVelocity;

END_FUNCTION

// Device/Application/02_Devices/F_Done
FUNCTION F_Done : BOOL
VAR_INPUT
    stStatus : ST_DeviceStatus;
    udiID : UDINT;
END_VAR

F_Done := (udiID <> 0) AND (stStatus.udiCompletedID = udiID)
    AND NOT stStatus.xBusy AND NOT stStatus.xError;

END_FUNCTION

// Device/Application/04_Machine/FB_AutoCycle
FUNCTION_BLOCK FB_AutoCycle
VAR_INPUT
    xRun : BOOL;
    xContinuous : BOOL;
    xMaterialAtLength : BOOL;
    stRecipe : ST_Recipe;
END_VAR
VAR_IN_OUT
    aCommand : ARRAY[1..17] OF ST_DeviceCommand;
    aStatus : ARRAY[1..17] OF ST_DeviceStatus;
    udiCounter : UDINT;
END_VAR
VAR_OUTPUT
    eStep : E_AutoStep;
    xDone : BOOL;
    xError : BOOL;
    udiErrorID : UDINT;
    uiClearLengthStep : UINT;
    uiClearTransferStep : UINT;
    uiPostStep : UINT;
    uiReturnKnifeStep : UINT;
    uiUnloadStep : UINT;
    uiResetLengthStep : UINT;
END_VAR
VAR
    ePrevStep : E_AutoStep := E_AutoStep.Fault;
    udiToken : UDINT;
    udiSpindleToken : UDINT;
    xEntry : BOOL;
    xSawSensorClear : BOOL;
    tonStep : TON;
    fbClear : FB_ClearanceUnit;
    fbPost : FB_PostCut;
END_VAR

xDone := FALSE;
IF NOT xRun THEN eStep:=E_AutoStep.Idle; xError:=FALSE; udiErrorID:=0; xSawSensorClear:=FALSE; END_IF
xEntry := eStep <> ePrevStep;
IF xEntry THEN udiToken := F_NextID(udiCounter); END_IF
ePrevStep := eStep;
tonStep(IN:=xRun AND NOT xEntry AND (eStep<>E_AutoStep.Idle)
    AND (eStep<>E_AutoStep.FeedWait) AND (eStep<>E_AutoStep.Complete)
    AND (eStep<>E_AutoStep.Fault),PT:=stRecipe.tStepTimeout);
IF xRun AND NOT xError THEN
CASE eStep OF
E_AutoStep.Idle: eStep:=E_AutoStep.FeedWait;
E_AutoStep.FeedWait:
    IF xEntry THEN xSawSensorClear:=FALSE; END_IF
    IF NOT xMaterialAtLength THEN xSawSensorClear:=TRUE; END_IF
    aCommand[1]:=F_Command(E_DeviceAction.Run,udiToken,0.0,stRecipe.lrBeltVelocity);
    IF xSawSensorClear AND xMaterialAtLength AND F_At(aStatus[5],1.0) THEN eStep:=E_AutoStep.StopFeed; END_IF
E_AutoStep.StopFeed:
    IF NOT aStatus[1].xActive AND NOT aStatus[1].xBusy THEN eStep:=E_AutoStep.Push; END_IF
E_AutoStep.Push:
    aCommand[11]:=F_Command(E_DeviceAction.Position,udiToken,1.0,stRecipe.lrPositionVelocity);
    IF F_Done(aStatus[11],udiToken) THEN eStep:=E_AutoStep.Clearance; END_IF
E_AutoStep.Clearance:
    IF fbClear.xDone THEN eStep:=E_AutoStep.Rotate; END_IF
E_AutoStep.Rotate:
    aCommand[8]:=F_Command(E_DeviceAction.Position,udiToken,stRecipe.lrRotateAngle,stRecipe.lrPositionVelocity);
    IF F_Done(aStatus[8],udiToken) THEN eStep:=E_AutoStep.PressDown; END_IF
E_AutoStep.PressDown:
    aCommand[9]:=F_Command(E_DeviceAction.Position,udiToken,1.0,stRecipe.lrPositionVelocity);
    IF F_Done(aStatus[9],udiToken) THEN eStep:=E_AutoStep.KnifeDown; END_IF
E_AutoStep.KnifeDown:
    aCommand[17]:=F_Command(E_DeviceAction.Position,udiToken,1.0,stRecipe.lrPositionVelocity);
    IF F_Done(aStatus[17],udiToken) THEN eStep:=E_AutoStep.SpindleOn; END_IF
E_AutoStep.SpindleOn:
    udiSpindleToken:=udiToken;
    aCommand[3]:=F_Command(E_DeviceAction.Run,udiSpindleToken,0.0,stRecipe.lrSpindleVelocity);
    IF F_Done(aStatus[3],udiSpindleToken) AND aStatus[3].xActive THEN eStep:=E_AutoStep.Cutting; END_IF
E_AutoStep.Cutting:
    aCommand[3]:=F_Command(E_DeviceAction.Run,udiSpindleToken,0.0,stRecipe.lrSpindleVelocity);
    aCommand[14]:=F_Command(E_DeviceAction.Run,udiToken,0.0,0.0);
    aCommand[2]:=F_Command(E_DeviceAction.Position,udiToken,stRecipe.lrCutHome+stRecipe.lrCutLength,stRecipe.lrCutVelocity);
    IF F_Done(aStatus[2],udiToken) THEN eStep:=E_AutoStep.StopCut; END_IF
E_AutoStep.StopCut:
    IF NOT aStatus[3].xActive AND NOT aStatus[3].xBusy AND NOT aStatus[14].xActive THEN eStep:=E_AutoStep.PostCut; END_IF
E_AutoStep.PostCut:
    IF fbPost.xDone THEN eStep:=E_AutoStep.Complete; END_IF
E_AutoStep.Complete:
    xDone:=xEntry;
    IF xContinuous THEN eStep:=E_AutoStep.FeedWait; END_IF
E_AutoStep.Fault: xError:=TRUE;
ELSE xError:=TRUE; udiErrorID:=4800;
END_CASE
IF tonStep.Q THEN xError:=TRUE; udiErrorID:=4800+TO_UDINT(eStep); END_IF
END_IF
fbClear(xExecute:=xRun AND (eStep=E_AutoStep.Clearance),stRecipe:=stRecipe,aCommand:=aCommand,aStatus:=aStatus,udiCounter:=udiCounter);
fbPost(xExecute:=xRun AND (eStep=E_AutoStep.PostCut),stRecipe:=stRecipe,aCommand:=aCommand,aStatus:=aStatus,udiCounter:=udiCounter);
IF fbClear.xError OR fbPost.xError THEN xError:=TRUE; udiErrorID:=MAX(fbClear.udiErrorID,fbPost.udiErrorID); END_IF
IF xError THEN eStep:=E_AutoStep.Fault; END_IF
uiClearLengthStep:=fbClear.uiLengthStep; uiClearTransferStep:=fbClear.uiTransferStep;
uiPostStep:=fbPost.uiStep; uiReturnKnifeStep:=fbPost.uiKnifeStep;
uiUnloadStep:=fbPost.uiUnloadStep; uiResetLengthStep:=fbPost.uiLengthStep;

END_FUNCTION_BLOCK

// Device/Application/02_Devices/F_At
FUNCTION F_At : BOOL
VAR_INPUT
    stStatus : ST_DeviceStatus;
    lrTarget : LREAL;
END_VAR

F_At := stStatus.xReady AND NOT stStatus.xBusy
    AND NOT stStatus.xError AND (ABS(stStatus.lrPosition-lrTarget) < 0.01);

END_FUNCTION

// Device/Application/03_Units/FB_ClearanceUnit
FUNCTION_BLOCK FB_ClearanceUnit
VAR_INPUT
    xExecute : BOOL;
    stRecipe : ST_Recipe;
END_VAR
VAR_IN_OUT
    aCommand : ARRAY[1..17] OF ST_DeviceCommand;
    aStatus : ARRAY[1..17] OF ST_DeviceStatus;
    udiCounter : UDINT;
END_VAR
VAR_OUTPUT
    xDone : BOOL;
    xError : BOOL;
    udiErrorID : UDINT;
    uiLengthStep : UINT;
    uiTransferStep : UINT;
END_VAR
VAR
    fbLength : FB_ClearLength;
    fbTransfer : FB_ClearTransfer;
END_VAR

fbLength(xExecute:=xExecute,stRecipe:=stRecipe,aCommand:=aCommand,aStatus:=aStatus,udiCounter:=udiCounter);
fbTransfer(xExecute:=xExecute,stRecipe:=stRecipe,aCommand:=aCommand,aStatus:=aStatus,udiCounter:=udiCounter);
xDone := fbLength.xDone AND fbTransfer.xDone;
xError := fbLength.xError OR fbTransfer.xError;
udiErrorID := MAX(fbLength.udiErrorID,fbTransfer.udiErrorID);
uiLengthStep := fbLength.uiStep; uiTransferStep := fbTransfer.uiStep;

END_FUNCTION_BLOCK

// Device/Application/03_Units/FB_ClearLength
FUNCTION_BLOCK FB_ClearLength
VAR_INPUT
    xExecute : BOOL;
    stRecipe : ST_Recipe;
END_VAR
VAR_IN_OUT
    aCommand : ARRAY[1..17] OF ST_DeviceCommand;
    aStatus : ARRAY[1..17] OF ST_DeviceStatus;
    udiCounter : UDINT;
END_VAR
VAR_OUTPUT
    xDone : BOOL;
    xError : BOOL;
    udiErrorID : UDINT;
    uiStep : UINT;
END_VAR
VAR
    uiPrevStep : UINT := 65535;
    udiToken : UDINT;
    xEntry : BOOL;
    tonStep : TON;
    tonSpray : TON;
END_VAR

IF NOT xExecute THEN uiStep := 0; xError := FALSE; udiErrorID := 0; END_IF;
xEntry := uiStep <> uiPrevStep;
IF xEntry THEN udiToken := F_NextID(udiCounter); END_IF;
uiPrevStep := uiStep;
tonStep(IN := xExecute AND (uiStep > 0) AND (uiStep < 1000) AND NOT xEntry, PT := stRecipe.tStepTimeout);
tonSpray(IN := xExecute AND (uiStep = 10) AND aStatus[13].xActive, PT := stRecipe.tSpray);
IF xExecute AND NOT xError THEN
CASE uiStep OF
0: uiStep := 10;
10: (* P010 length up *)
aCommand[5] := F_Command(E_DeviceAction.Position, udiToken, 0.0, stRecipe.lrPositionVelocity);
IF F_Done(aStatus[5], udiToken) THEN uiStep := 20; END_IF;
20: (* P020 move length clear *)
aCommand[4] := F_Command(E_DeviceAction.Position, udiToken, stRecipe.lrLengthClear, stRecipe.lrPositionVelocity);
IF F_Done(aStatus[4], udiToken) THEN uiStep := 1000; END_IF;
1000: ;
ELSE xError := TRUE; udiErrorID := 4100;
END_CASE;
IF tonStep.Q THEN xError := TRUE; udiErrorID := 4100 + UINT_TO_UDINT(uiStep); END_IF;
END_IF;
xDone := xExecute AND (uiStep = 1000) AND NOT xError;

END_FUNCTION_BLOCK

// Device/Application/03_Units/FB_ClearTransfer
FUNCTION_BLOCK FB_ClearTransfer
VAR_INPUT
    xExecute : BOOL;
    stRecipe : ST_Recipe;
END_VAR
VAR_IN_OUT
    aCommand : ARRAY[1..17] OF ST_DeviceCommand;
    aStatus : ARRAY[1..17] OF ST_DeviceStatus;
    udiCounter : UDINT;
END_VAR
VAR_OUTPUT
    xDone : BOOL;
    xError : BOOL;
    udiErrorID : UDINT;
    uiStep : UINT;
END_VAR
VAR
    uiPrevStep : UINT := 65535;
    udiToken : UDINT;
    xEntry : BOOL;
    tonStep : TON;
    tonSpray : TON;
END_VAR

IF NOT xExecute THEN uiStep := 0; xError := FALSE; udiErrorID := 0; END_IF;
xEntry := uiStep <> uiPrevStep;
IF xEntry THEN udiToken := F_NextID(udiCounter); END_IF;
uiPrevStep := uiStep;
tonStep(IN := xExecute AND (uiStep > 0) AND (uiStep < 1000) AND NOT xEntry, PT := stRecipe.tStepTimeout);
tonSpray(IN := xExecute AND (uiStep = 10) AND aStatus[13].xActive, PT := stRecipe.tSpray);
IF xExecute AND NOT xError THEN
CASE uiStep OF
0: uiStep := 10;
10: (* Q010 roller down *)
aCommand[12] := F_Command(E_DeviceAction.Position, udiToken, 0.0, stRecipe.lrPositionVelocity);
IF F_Done(aStatus[12], udiToken) THEN uiStep := 20; END_IF;
20: (* Q020 release side push *)
aCommand[11] := F_Command(E_DeviceAction.Position, udiToken, 0.0, stRecipe.lrPositionVelocity);
IF F_Done(aStatus[11], udiToken) THEN uiStep := 30; END_IF;
30: (* Q030 lower selected side stop *)
aCommand[10] := F_Command(E_DeviceAction.Position, udiToken, 1.0, stRecipe.lrPositionVelocity);
IF F_Done(aStatus[10], udiToken) THEN uiStep := 1000; END_IF;
1000: ;
ELSE xError := TRUE; udiErrorID := 4200;
END_CASE;
IF tonStep.Q THEN xError := TRUE; udiErrorID := 4200 + UINT_TO_UDINT(uiStep); END_IF;
END_IF;
xDone := xExecute AND (uiStep = 1000) AND NOT xError;

END_FUNCTION_BLOCK

// Device/Application/03_Units/FB_PostCut
FUNCTION_BLOCK FB_PostCut
VAR_INPUT
    xExecute : BOOL;
    stRecipe : ST_Recipe;
END_VAR
VAR_IN_OUT
    aCommand : ARRAY[1..17] OF ST_DeviceCommand;
    aStatus : ARRAY[1..17] OF ST_DeviceStatus;
    udiCounter : UDINT;
END_VAR
VAR_OUTPUT
    xDone : BOOL;
    xError : BOOL;
    udiErrorID : UDINT;
    uiStep : UINT;
    uiKnifeStep : UINT;
    uiUnloadStep : UINT;
    uiLengthStep : UINT;
END_VAR
VAR
    fbKnife : FB_ReturnKnife;
    fbUnload : FB_Unload;
    fbLength : FB_ResetLength;
    uiPrevStep : UINT := 65535;
    udiToken : UDINT;
    xEntry : BOOL;
    tonStep : TON;
END_VAR

IF NOT xExecute THEN uiStep := 0; xError := FALSE; udiErrorID := 0; END_IF
xEntry := uiStep <> uiPrevStep;
IF xEntry THEN udiToken := F_NextID(udiCounter); END_IF
uiPrevStep := uiStep;
tonStep(IN:=xExecute AND NOT xEntry AND (uiStep>0) AND (uiStep<1000),PT:=stRecipe.tStepTimeout);
IF xExecute AND NOT xError THEN
    CASE uiStep OF
    0: uiStep := 10;
    10:
        aCommand[17] := F_Command(E_DeviceAction.Position,udiToken,0.0,stRecipe.lrPositionVelocity);
        IF F_Done(aStatus[17],udiToken) THEN uiStep := 20; END_IF
    20:
        aCommand[9] := F_Command(E_DeviceAction.Position,udiToken,0.0,stRecipe.lrPositionVelocity);
        IF F_Done(aStatus[9],udiToken) THEN uiStep := 30; END_IF
    30:
        IF fbKnife.xDone AND fbUnload.xDone AND fbLength.xDone THEN uiStep := 1000; END_IF
    1000: ;
    ELSE xError := TRUE; udiErrorID := 4700;
    END_CASE
    IF tonStep.Q THEN xError := TRUE; udiErrorID := 4700+UINT_TO_UDINT(uiStep); END_IF
END_IF
fbKnife(xExecute:=xExecute AND (uiStep=30),stRecipe:=stRecipe,aCommand:=aCommand,aStatus:=aStatus,udiCounter:=udiCounter);
fbUnload(xExecute:=xExecute AND (uiStep=30),stRecipe:=stRecipe,aCommand:=aCommand,aStatus:=aStatus,udiCounter:=udiCounter);
fbLength(xExecute:=xExecute AND (uiStep=30),stRecipe:=stRecipe,aCommand:=aCommand,aStatus:=aStatus,udiCounter:=udiCounter);
IF fbKnife.xError OR fbUnload.xError OR fbLength.xError THEN
    xError:=TRUE; udiErrorID:=MAX(fbKnife.udiErrorID,MAX(fbUnload.udiErrorID,fbLength.udiErrorID));
END_IF
xDone := xExecute AND (uiStep=1000) AND NOT xError;
uiKnifeStep:=fbKnife.uiStep; uiUnloadStep:=fbUnload.uiStep; uiLengthStep:=fbLength.uiStep;

END_FUNCTION_BLOCK

// Device/Application/03_Units/FB_ReturnKnife
FUNCTION_BLOCK FB_ReturnKnife
VAR_INPUT
    xExecute : BOOL;
    stRecipe : ST_Recipe;
END_VAR
VAR_IN_OUT
    aCommand : ARRAY[1..17] OF ST_DeviceCommand;
    aStatus : ARRAY[1..17] OF ST_DeviceStatus;
    udiCounter : UDINT;
END_VAR
VAR_OUTPUT
    xDone : BOOL;
    xError : BOOL;
    udiErrorID : UDINT;
    uiStep : UINT;
END_VAR
VAR
    uiPrevStep : UINT := 65535;
    udiToken : UDINT;
    xEntry : BOOL;
    tonStep : TON;
    tonSpray : TON;
END_VAR

IF NOT xExecute THEN uiStep := 0; xError := FALSE; udiErrorID := 0; END_IF;
xEntry := uiStep <> uiPrevStep;
IF xEntry THEN udiToken := F_NextID(udiCounter); END_IF;
uiPrevStep := uiStep;
tonStep(IN := xExecute AND (uiStep > 0) AND (uiStep < 1000) AND NOT xEntry, PT := stRecipe.tStepTimeout);
tonSpray(IN := xExecute AND (uiStep = 10) AND aStatus[13].xActive, PT := stRecipe.tSpray);
IF xExecute AND NOT xError THEN
CASE uiStep OF
0: uiStep := 10;
10: (* A010 spray before return *)
aCommand[13] := F_Command(E_DeviceAction.Run, udiToken, 0.0, 0.0);
IF tonSpray.Q THEN uiStep := 20; END_IF;
20: (* A020 return cut axis *)
aCommand[2] := F_Command(E_DeviceAction.Position, udiToken, stRecipe.lrCutHome, stRecipe.lrPositionVelocity);
IF F_Done(aStatus[2], udiToken) THEN uiStep := 1000; END_IF;
1000: ;
ELSE xError := TRUE; udiErrorID := 4300;
END_CASE;
IF tonStep.Q THEN xError := TRUE; udiErrorID := 4300 + UINT_TO_UDINT(uiStep); END_IF;
END_IF;
xDone := xExecute AND (uiStep = 1000) AND NOT xError;

END_FUNCTION_BLOCK

// Device/Application/03_Units/FB_Unload
FUNCTION_BLOCK FB_Unload
VAR_INPUT
    xExecute : BOOL;
    stRecipe : ST_Recipe;
END_VAR
VAR_IN_OUT
    aCommand : ARRAY[1..17] OF ST_DeviceCommand;
    aStatus : ARRAY[1..17] OF ST_DeviceStatus;
    udiCounter : UDINT;
END_VAR
VAR_OUTPUT
    xDone : BOOL;
    xError : BOOL;
    udiErrorID : UDINT;
    uiStep : UINT;
END_VAR
VAR
    uiPrevStep : UINT := 65535;
    udiToken : UDINT;
    xEntry : BOOL;
    tonStep : TON;
    tonSpray : TON;
END_VAR

IF NOT xExecute THEN uiStep := 0; xError := FALSE; udiErrorID := 0; END_IF;
xEntry := uiStep <> uiPrevStep;
IF xEntry THEN udiToken := F_NextID(udiCounter); END_IF;
uiPrevStep := uiStep;
tonStep(IN := xExecute AND (uiStep > 0) AND (uiStep < 1000) AND NOT xEntry, PT := stRecipe.tStepTimeout);
tonSpray(IN := xExecute AND (uiStep = 10) AND aStatus[13].xActive, PT := stRecipe.tSpray);
IF xExecute AND NOT xError THEN
CASE uiStep OF
0: uiStep := 10;
10: (* B010 side stop up *)
aCommand[10] := F_Command(E_DeviceAction.Position, udiToken, 0.0, stRecipe.lrPositionVelocity);
IF F_Done(aStatus[10], udiToken) THEN uiStep := 20; END_IF;
20: (* B020 rollers up *)
aCommand[12] := F_Command(E_DeviceAction.Position, udiToken, 1.0, stRecipe.lrPositionVelocity);
IF F_Done(aStatus[12], udiToken) THEN uiStep := 30; END_IF;
30: (* B030 gripper lift up *)
aCommand[15] := F_Command(E_DeviceAction.Position, udiToken, 1.0, stRecipe.lrPositionVelocity);
IF F_Done(aStatus[15], udiToken) THEN uiStep := 40; END_IF;
40: (* B040 gripper open *)
aCommand[16] := F_Command(E_DeviceAction.Position, udiToken, 0.0, stRecipe.lrPositionVelocity);
IF F_Done(aStatus[16], udiToken) THEN uiStep := 50; END_IF;
50: (* B050 gripper forward *)
aCommand[7] := F_Command(E_DeviceAction.Position, udiToken, stRecipe.lrGripperFront, stRecipe.lrPositionVelocity);
IF F_Done(aStatus[7], udiToken) THEN uiStep := 60; END_IF;
60: (* B060 gripper clamp *)
aCommand[16] := F_Command(E_DeviceAction.Position, udiToken, 1.0, stRecipe.lrPositionVelocity);
IF F_Done(aStatus[16], udiToken) THEN uiStep := 70; END_IF;
70: (* B070 pull product *)
aCommand[7] := F_Command(E_DeviceAction.Position, udiToken, stRecipe.lrGripperPull, stRecipe.lrPositionVelocity);
IF F_Done(aStatus[7], udiToken) THEN uiStep := 80; END_IF;
80: (* B080 gripper open *)
aCommand[16] := F_Command(E_DeviceAction.Position, udiToken, 0.0, stRecipe.lrPositionVelocity);
IF F_Done(aStatus[16], udiToken) THEN uiStep := 90; END_IF;
90: (* B090 retreat while raised *)
aCommand[7] := F_Command(E_DeviceAction.Position, udiToken, stRecipe.lrGripperBack, stRecipe.lrPositionVelocity);
IF F_Done(aStatus[7], udiToken) THEN uiStep := 100; END_IF;
100: (* B100 lower gripper *)
aCommand[15] := F_Command(E_DeviceAction.Position, udiToken, 0.0, stRecipe.lrPositionVelocity);
IF F_Done(aStatus[15], udiToken) THEN uiStep := 110; END_IF;
110: (* B110 final return while lowered *)
aCommand[7] := F_Command(E_DeviceAction.Position, udiToken, stRecipe.lrGripperHome, stRecipe.lrPositionVelocity);
IF F_Done(aStatus[7], udiToken) THEN uiStep := 1000; END_IF;
1000: ;
ELSE xError := TRUE; udiErrorID := 4400;
END_CASE;
IF tonStep.Q THEN xError := TRUE; udiErrorID := 4400 + UINT_TO_UDINT(uiStep); END_IF;
END_IF;
xDone := xExecute AND (uiStep = 1000) AND NOT xError;

END_FUNCTION_BLOCK

// Device/Application/03_Units/FB_ResetLength
FUNCTION_BLOCK FB_ResetLength
VAR_INPUT
    xExecute : BOOL;
    stRecipe : ST_Recipe;
END_VAR
VAR_IN_OUT
    aCommand : ARRAY[1..17] OF ST_DeviceCommand;
    aStatus : ARRAY[1..17] OF ST_DeviceStatus;
    udiCounter : UDINT;
END_VAR
VAR_OUTPUT
    xDone : BOOL;
    xError : BOOL;
    udiErrorID : UDINT;
    uiStep : UINT;
END_VAR
VAR
    uiPrevStep : UINT := 65535;
    udiToken : UDINT;
    xEntry : BOOL;
    tonStep : TON;
    tonSpray : TON;
END_VAR

IF NOT xExecute THEN uiStep := 0; xError := FALSE; udiErrorID := 0; END_IF;
xEntry := uiStep <> uiPrevStep;
IF xEntry THEN udiToken := F_NextID(udiCounter); END_IF;
uiPrevStep := uiStep;
tonStep(IN := xExecute AND (uiStep > 0) AND (uiStep < 1000) AND NOT xEntry, PT := stRecipe.tStepTimeout);
tonSpray(IN := xExecute AND (uiStep = 10) AND aStatus[13].xActive, PT := stRecipe.tSpray);
IF xExecute AND NOT xError THEN
CASE uiStep OF
0: uiStep := 10;
10: (* C010 length to detection position *)
aCommand[4] := F_Command(E_DeviceAction.Position, udiToken, stRecipe.lrLengthPosition, stRecipe.lrPositionVelocity);
IF F_Done(aStatus[4], udiToken) THEN uiStep := 20; END_IF;
20: (* C020 lower length sensor *)
aCommand[5] := F_Command(E_DeviceAction.Position, udiToken, 1.0, stRecipe.lrPositionVelocity);
IF F_Done(aStatus[5], udiToken) THEN uiStep := 30; END_IF;
30: (* C030 verify down, detection permission follows physical position *)
IF F_At(aStatus[5],1.0) THEN uiStep := 1000; END_IF;
1000: ;
ELSE xError := TRUE; udiErrorID := 4500;
END_CASE;
IF tonStep.Q THEN xError := TRUE; udiErrorID := 4500 + UINT_TO_UDINT(uiStep); END_IF;
END_IF;
xDone := xExecute AND (uiStep = 1000) AND NOT xError;

END_FUNCTION_BLOCK

// Device/Application/03_Units/FB_Initialize
FUNCTION_BLOCK FB_Initialize
VAR_INPUT
    xExecute : BOOL;
    stRecipe : ST_Recipe;
END_VAR
VAR_IN_OUT
    aCommand : ARRAY[1..17] OF ST_DeviceCommand;
    aStatus : ARRAY[1..17] OF ST_DeviceStatus;
    udiCounter : UDINT;
END_VAR
VAR_OUTPUT
    xDone : BOOL;
    xError : BOOL;
    udiErrorID : UDINT;
    uiStep : UINT;
END_VAR
VAR
    uiPrevStep : UINT := 65535;
    udiToken : UDINT;
    xEntry : BOOL;
    tonStep : TON;
    tonSpray : TON;
END_VAR

IF NOT xExecute THEN uiStep := 0; xError := FALSE; udiErrorID := 0; END_IF;
xEntry := uiStep <> uiPrevStep;
IF xEntry THEN udiToken := F_NextID(udiCounter); END_IF;
uiPrevStep := uiStep;
tonStep(IN := xExecute AND (uiStep > 0) AND (uiStep < 1000) AND NOT xEntry, PT := stRecipe.tStepTimeout);
tonSpray(IN := xExecute AND (uiStep = 10) AND aStatus[13].xActive, PT := stRecipe.tSpray);
IF xExecute AND NOT xError THEN
CASE uiStep OF
0: uiStep := 10;
10: (* SIMULATION initialization: lift knife, press; open gripper *)
aCommand[17] := F_Command(E_DeviceAction.Position, udiToken, 0.0, stRecipe.lrPositionVelocity);
aCommand[9] := F_Command(E_DeviceAction.Position, udiToken, 0.0, stRecipe.lrPositionVelocity);
aCommand[16] := F_Command(E_DeviceAction.Position, udiToken, 0.0, stRecipe.lrPositionVelocity);
IF F_Done(aStatus[17], udiToken) AND F_Done(aStatus[9], udiToken) AND F_Done(aStatus[16], udiToken) THEN uiStep := 20; END_IF;
20: (* Prepare clear positions *)
aCommand[5] := F_Command(E_DeviceAction.Position, udiToken, 0.0, stRecipe.lrPositionVelocity);
aCommand[10] := F_Command(E_DeviceAction.Position, udiToken, 0.0, stRecipe.lrPositionVelocity);
aCommand[11] := F_Command(E_DeviceAction.Position, udiToken, 0.0, stRecipe.lrPositionVelocity);
aCommand[12] := F_Command(E_DeviceAction.Position, udiToken, 1.0, stRecipe.lrPositionVelocity);
aCommand[15] := F_Command(E_DeviceAction.Position, udiToken, 0.0, stRecipe.lrPositionVelocity);
IF F_Done(aStatus[5], udiToken) AND F_Done(aStatus[10], udiToken) AND F_Done(aStatus[11], udiToken) AND F_Done(aStatus[12], udiToken) AND F_Done(aStatus[15], udiToken) THEN uiStep := 30; END_IF;
30: (* Move to simulation initial coordinates *)
aCommand[2] := F_Command(E_DeviceAction.Position, udiToken, stRecipe.lrCutHome, stRecipe.lrPositionVelocity);
aCommand[4] := F_Command(E_DeviceAction.Position, udiToken, stRecipe.lrLengthPosition, stRecipe.lrPositionVelocity);
aCommand[7] := F_Command(E_DeviceAction.Position, udiToken, stRecipe.lrGripperHome, stRecipe.lrPositionVelocity);
aCommand[8] := F_Command(E_DeviceAction.Position, udiToken, 0.0, stRecipe.lrPositionVelocity);
IF F_Done(aStatus[2], udiToken) AND F_Done(aStatus[4], udiToken) AND F_Done(aStatus[7], udiToken) AND F_Done(aStatus[8], udiToken) THEN uiStep := 40; END_IF;
40: (* Length down for detection *)
aCommand[5] := F_Command(E_DeviceAction.Position, udiToken, 1.0, stRecipe.lrPositionVelocity);
IF F_Done(aStatus[5], udiToken) THEN uiStep := 1000; END_IF;
1000: ;
ELSE xError := TRUE; udiErrorID := 4600;
END_CASE;
IF tonStep.Q THEN xError := TRUE; udiErrorID := 4600 + UINT_TO_UDINT(uiStep); END_IF;
END_IF;
xDone := xExecute AND (uiStep = 1000) AND NOT xError;

END_FUNCTION_BLOCK

// Device/Application/04_Machine/FB_Interlocks
FUNCTION_BLOCK FB_Interlocks
VAR_INPUT
    xPermit : BOOL;
    stRecipe : ST_Recipe;
    aRequest : ARRAY[1..17] OF ST_DeviceCommand;
    aStatus : ARRAY[1..17] OF ST_DeviceStatus;
END_VAR
VAR_OUTPUT
    aCommand : ARRAY[1..17] OF ST_DeviceCommand;
    uiBlockedDevice : UINT;
END_VAR
VAR
    i : INT;
    xAllowed : BOOL;
    xMotion : BOOL;
    xKnifeUp : BOOL;
    xPressUp : BOOL;
    xClampOpen : BOOL;
END_VAR

uiBlockedDevice:=0;
xKnifeUp:=F_At(aStatus[17],0.0); xPressUp:=F_At(aStatus[9],0.0);
xClampOpen:=F_At(aStatus[16],0.0);
FOR i:=1 TO 17 DO
    aCommand[i]:=aRequest[i];
    xAllowed:=xPermit AND (i<>6);
    xMotion:=(aRequest[i].eAction=E_DeviceAction.Jog) OR
        ((aRequest[i].eAction=E_DeviceAction.Position) AND
        (ABS(aRequest[i].lrTarget-aStatus[i].lrPosition)>0.01));
    IF xMotion THEN
        CASE i OF
        4: xAllowed:=xAllowed AND F_At(aStatus[5],0.0);
        8: xAllowed:=xAllowed AND xKnifeUp AND xPressUp AND F_At(aStatus[11],0.0);
        9:
            IF aRequest[i].lrTarget>0.5 THEN
                xAllowed:=xAllowed AND NOT aStatus[8].xBusy AND xKnifeUp AND F_At(aStatus[2],stRecipe.lrCutHome);
            END_IF
        17:
            IF aRequest[i].lrTarget>0.5 THEN
                xAllowed:=xAllowed AND F_At(aStatus[9],1.0) AND NOT aStatus[8].xBusy
                    AND F_At(aStatus[5],0.0) AND F_At(aStatus[12],0.0) AND F_At(aStatus[10],1.0);
            END_IF
        2:
            IF ((aRequest[i].eAction=E_DeviceAction.Position) AND (aRequest[i].lrTarget>stRecipe.lrCutHome+0.01))
               OR ((aRequest[i].eAction=E_DeviceAction.Jog) AND (aRequest[i].lrVelocity>0.0)) THEN
                xAllowed:=xAllowed AND F_At(aStatus[9],1.0) AND F_At(aStatus[17],1.0) AND aStatus[3].xActive;
            ELSE xAllowed:=xAllowed AND xKnifeUp;
            END_IF
        7:
            xAllowed:=xAllowed AND xKnifeUp AND xPressUp;
            IF aRequest[i].eAction=E_DeviceAction.Jog THEN
                xAllowed:=xAllowed AND F_At(aStatus[15],1.0) AND xClampOpen;
            ELSIF ABS(aRequest[i].lrTarget-stRecipe.lrGripperHome)<0.01 THEN
                xAllowed:=xAllowed AND F_At(aStatus[15],0.0) AND xClampOpen;
            ELSIF ABS(aRequest[i].lrTarget-stRecipe.lrGripperPull)<0.01 THEN
                xAllowed:=xAllowed AND F_At(aStatus[15],1.0) AND F_At(aStatus[16],1.0);
            ELSE xAllowed:=xAllowed AND F_At(aStatus[15],1.0) AND xClampOpen;
            END_IF
        END_CASE
    END_IF
    IF NOT xAllowed THEN
        IF aRequest[i].eAction<>E_DeviceAction.None THEN uiBlockedDevice:=INT_TO_UINT(i); END_IF
        aCommand[i].eAction:=E_DeviceAction.Stop;
    END_IF
END_FOR

END_FUNCTION_BLOCK

// Device/Application/06_Simulation/FB_SimPlant
FUNCTION_BLOCK FB_SimPlant
VAR_INPUT
    xEnable : BOOL;
    stSettings : ST_SimulationSettings;
    aStatus : ARRAY[1..17] OF ST_DeviceStatus;
END_VAR
VAR_OUTPUT
    xMaterialAtLength : BOOL;
END_VAR
VAR
    xLatched : BOOL;
    tonMaterial : TON;
END_VAR

IF NOT xEnable OR NOT F_At(aStatus[5],1.0) THEN xLatched:=FALSE; END_IF
tonMaterial(IN:=xEnable AND stSettings.xAutoMaterial AND aStatus[1].xActive
    AND F_At(aStatus[5],1.0) AND NOT xLatched,PT:=stSettings.tMaterialDelay);
IF tonMaterial.Q THEN xLatched:=TRUE; END_IF
IF stSettings.xAutoMaterial THEN xMaterialAtLength:=xLatched;
ELSE xMaterialAtLength:=xEnable AND F_At(aStatus[5],1.0) AND stSettings.xMaterialSensor;
END_IF

END_FUNCTION_BLOCK

// Device/Application/04_Machine/FB_AlarmManager
FUNCTION_BLOCK FB_AlarmManager
VAR_INPUT
    udiIncoming : UDINT;
    xReset : BOOL;
END_VAR
VAR_OUTPUT
    udiLatched : UDINT;
END_VAR

IF xReset AND (udiIncoming=0) THEN udiLatched:=0; END_IF
IF (udiLatched=0) AND (udiIncoming<>0) THEN udiLatched:=udiIncoming; END_IF

END_FUNCTION_BLOCK

// Device/Application/04_Machine/FB_IOMap
FUNCTION_BLOCK FB_IOMap
VAR_INPUT
    uiMaterialModel : UINT;
    aCommand : ARRAY[1..17] OF ST_DeviceCommand;
    aStatus : ARRAY[1..17] OF ST_DeviceStatus;
END_VAR
VAR_IN_OUT
    axOutputs : ARRAY[0..31] OF BOOL;
    axG2RelayDemand : ARRAY[1..3] OF BOOL;
END_VAR
VAR
    i : INT;
END_VAR

(* Physical writes remain unimplemented. Logical relay demand is diagnostic. *)
FOR i:=0 TO 31 DO axOutputs[i]:=FALSE; END_FOR
FOR i:=1 TO 3 DO axG2RelayDemand[i]:=FALSE; END_FOR
IF aStatus[10].lrPosition>0.5 THEN
    CASE uiMaterialModel OF
    300: axG2RelayDemand[1]:=TRUE;
    400: axG2RelayDemand[2]:=TRUE;
    600: axG2RelayDemand[3]:=TRUE;
    END_CASE
END_IF

END_FUNCTION_BLOCK

// Device/Application/90_Legacy/PRG_AxisDemo
PROGRAM PRG_AxisDemo
VAR
    (* ---- SoftMotion function block instances ---- *)
    fbPower    : MC_Power;            (* enable / disable the axis *)
    fbReset    : MC_Reset;            (* reset axis error *)
    fbStop     : MC_Stop;             (* stop and lock the axis *)
    fbJog      : MC_Jog;              (* jog *)
    fbMoveRel  : MC_MoveRelative;     (* single relative move *)
    fbMoveAbs  : MC_MoveAbsolute;     (* single absolute move *)
    fbCycle    : MC_MoveRelative;     (* auto cycle move *)
    fbReadPos  : MC_ReadActualPosition; (* position feedback *)
    fbReadStat : MC_ReadStatus;       (* axis state machine *)
    fbReadErr  : MC_ReadAxisError;    (* axis error code *)

    (* ---- edge detection ---- *)
    rtCycle    : R_TRIG;              (* auto cycle trigger *)

    (* ---- auto cycle ---- *)
    fbCycleExec: BOOL;                (* Execute for fbCycle *)
    rCycleDist : LREAL;               (* current segment distance *)
    iCycle     : INT := 0;            (* auto cycle step *)
    tonDwell   : TON;                 (* dwell at cycle ends *)

    (* ---- diagnostics ---- *)
    eLastErr   : SMC_ERROR;           (* latched last motion block error *)
	xDoReset: BOOL;
	xStopRun: BOOL;
	rRunDec: LREAL;
	xStartRun: BOOL;
	iStep: INT;
	fbMoveVel: MC_MoveVelocity;
	Axis: INT;
	Execute: BOOL;
	rRunVel: LREAL;
	rRunAcc: LREAL;
	Velocity: INT;
	Acceleration: INT;
	Deceleration: INT;
	Direction: INT;
	InVelocity: INT;
	xMoveExec: BOOL;
END_VAR

(* Single low-speed 20 mm out-and-back test cycle.
   Start only on a rising edge of GVL_Motion.xStartCycle.
   Travel is capped at 20 mm per leg and 10 mm/s. *)
rtCycle(CLK := GVL_Motion.xStartCycle);

fbPower(Axis         := Axis_1,
        Enable       := GVL_Motion.xEnable,
        bRegulatorOn := TRUE,
        bDriveStart  := TRUE);

fbReset(Axis := Axis_1, Execute := GVL_Motion.xReset);

IF GVL_Motion.xStop THEN
    xStopRun   := TRUE;
    fbCycleExec := FALSE;
    iCycle      := 0;
END_IF

IF fbPower.Error OR fbCycle.Error OR fbReset.Error OR fbStop.Error THEN
    iCycle      := 99;
    fbCycleExec := FALSE;
    xStopRun    := TRUE;
END_IF

fbStop(Axis         := Axis_1,
       Execute      := xStopRun,
       Deceleration := MIN(MAX(GVL_Motion.rDec, 10.0), 200.0));

IF xStopRun AND fbStop.Done THEN
    xStopRun := FALSE;
END_IF

tonDwell(IN := (iCycle = 20) OR (iCycle = 40),
         PT := GVL_Motion.tDwell);

CASE iCycle OF
    0:  (* Idle; one rising edge starts one round trip. *)
        fbCycleExec := FALSE;
        IF rtCycle.Q
           AND GVL_Motion.xEnable
           AND fbPower.Status
           AND NOT GVL_Motion.xAxisError
           AND NOT xStopRun
           AND (ABS(GVL_Motion.rStroke) > 0.0) THEN
            rCycleDist := MIN(ABS(GVL_Motion.rStroke), 20.0);
            fbCycleExec := TRUE;
            iCycle := 10;
        END_IF

    10: (* Forward leg. *)
        IF fbCycle.Done THEN
            fbCycleExec := FALSE;
            iCycle := 20;
        ELSIF fbCycle.Error THEN
            fbCycleExec := FALSE;
            iCycle := 99;
            xStopRun := TRUE;
        END_IF

    20: (* Dwell before return leg. *)
        IF tonDwell.Q AND NOT xStopRun THEN
            rCycleDist := -MIN(ABS(GVL_Motion.rStroke), 20.0);
            fbCycleExec := TRUE;
            iCycle := 30;
        END_IF

    30: (* Return leg. *)
        IF fbCycle.Done THEN
            fbCycleExec := FALSE;
            iCycle := 40;
        ELSIF fbCycle.Error THEN
            fbCycleExec := FALSE;
            iCycle := 99;
            xStopRun := TRUE;
        END_IF

    40: (* Dwell after returning to the start position, then finish. *)
        IF tonDwell.Q THEN
            iCycle := 0;
        END_IF

    99: (* Error latch; require a successful reset and completed stop. *)
        fbCycleExec := FALSE;
        IF GVL_Motion.xReset AND fbReset.Done AND NOT xStopRun THEN
            iCycle := 0;
        END_IF

ELSE
    iCycle := 99;
    fbCycleExec := FALSE;
    xStopRun := TRUE;
END_CASE

fbCycle(Axis         := Axis_1,
        Execute      := fbCycleExec AND NOT xStopRun,
        Distance     := rCycleDist,
        Velocity     := MIN(MAX(GVL_Motion.rVel, 1.0), 10.0),
        Acceleration := MIN(MAX(GVL_Motion.rAcc, 10.0), 200.0),
        Deceleration := MIN(MAX(GVL_Motion.rDec, 10.0), 200.0));

fbReadPos(Axis := Axis_1, Enable := TRUE);

GVL_Motion.xPowered    := fbPower.Status;
GVL_Motion.xBusy       := fbCycle.Busy OR fbStop.Busy;
GVL_Motion.xDisabled   := NOT fbPower.Status;
GVL_Motion.xStopping   := fbStop.Busy;
GVL_Motion.xStandStill := fbPower.Status AND NOT GVL_Motion.xBusy;
GVL_Motion.xAxisReady  := GVL_Motion.xStandStill AND NOT GVL_Motion.xAxisError;
GVL_Motion.xAxisError  := fbPower.Error OR fbCycle.Error OR fbReset.Error OR fbStop.Error;
GVL_Motion.xErrorStop  := GVL_Motion.xAxisError;
GVL_Motion.iState      := iCycle;
GVL_Motion.rActPos     := fbReadPos.Position;

END_PROGRAM
